(* IEC 61131-3 sources: s7-to-codesys/tests/POUs/ScenariosLang/FB_ConveyorStl_ScenarioTest, 15 files *)

(* ---- FB_ConveyorStl_ScenarioTest.decl.st ---- *)
// AUTO-GENERATED — не редактировать: s7conv gen-tests, сценарии scenarios/lang/FB_ConveyorStl.csv
// Правка — в CSV (scenarios/README.md), затем python -m s7conv build-corpus.
// Назначение: тесты поведения сконвертированного FB_ConveyorStl по сценариям CSV (сценариев: 7, строк: 58):
//             один метод-тест на сценарий, строки — по порядку с моделируемым временем GVL_S7Clock.
//             Ожидаемые значения — из CSV (эталонные модели по описанию логики блока), не из
//             результата конвертации.
// Автор:      s7conv 0.1.0 (сгенерировано)
// Версия:     не указана
// Документ:   scenarios/README.md, docs/methodology.md, раздел «Проверка поведения»
FUNCTION_BLOCK FB_ConveyorStl_ScenarioTest EXTENDS coUnit.FB_TestSuite
VAR
    fbStartSequence : FB_ConveyorStl;  // свой экземпляр на сценарий
    xStartSequenceDone : BOOL;  // сценарий выполнен (выполняется один раз)
    fbStopRunOut : FB_ConveyorStl;  // свой экземпляр на сценарий
    xStopRunOutDone : BOOL;  // сценарий выполнен (выполняется один раз)
    fbJamWithoutProducts : FB_ConveyorStl;  // свой экземпляр на сценарий
    xJamWithoutProductsDone : BOOL;  // сценарий выполнен (выполняется один раз)
    fbProductsKeepFlow : FB_ConveyorStl;  // свой экземпляр на сценарий
    xProductsKeepFlowDone : BOOL;  // сценарий выполнен (выполняется один раз)
    fbCountResetIsLevel : FB_ConveyorStl;  // свой экземпляр на сценарий
    xCountResetIsLevelDone : BOOL;  // сценарий выполнен (выполняется один раз)
    fbHornCutShort : FB_ConveyorStl;  // свой экземпляр на сценарий
    xHornCutShortDone : BOOL;  // сценарий выполнен (выполняется один раз)
    fbAckRestartsFlowWatch : FB_ConveyorStl;  // свой экземпляр на сценарий
    xAckRestartsFlowWatchDone : BOOL;  // сценарий выполнен (выполняется один раз)
END_VAR

(* ---- AckRestartsFlowWatch.method.decl.st ---- *)
// AUTO-GENERATED — не редактировать: scenarios/lang/FB_ConveyorStl.csv, сценарий AckRestartsFlowWatch (строк: 10)
METHOD PRIVATE AckRestartsFlowWatch
VAR
    stTimerZero : ST_S5Timer;  // пустое слово S5 для сброса
    stCounterZero : ST_S5Counter;  // пустое слово S5 для сброса
    iS5 : INT;  // номер таймера/счётчика S5
END_VAR

(* ---- AckRestartsFlowWatch.method.impl.st ---- *)
// AUTO-GENERATED — не редактировать: scenarios/lang/FB_ConveyorStl.csv, сценарий AckRestartsFlowWatch
coUnit.TEST('AckRestartsFlowWatch');
IF NOT xAckRestartsFlowWatchDone THEN
    xAckRestartsFlowWatchDone := TRUE;
    GVL_S7Clock.xSimulation := TRUE;
    // слова S5 — глобальные (GVL_S5Timers_Lang): сценарий начинается с чистых таймеров и счётчиков
    FOR iS5 := 0 TO 5 DO
        GVL_S5Timers_Lang.aTimer[iS5] := stTimerZero;
    END_FOR
    // слова S5 — глобальные (GVL_S5Counters_Lang): сценарий начинается с чистых таймеров и счётчиков
    FOR iS5 := 0 TO 1 DO
        GVL_S5Counters_Lang.aCounter[iS5] := stCounterZero;
    END_FOR

    // #1, t = 0 мс — пуск: запрос, сирена T1 и задержка T2 пошли
    GVL_S7Clock.tSimNow := T#0MS;
    fbAckRestartsFlowWatch.xStart := TRUE;
    fbAckRestartsFlowWatch.xStop := FALSE;
    fbAckRestartsFlowWatch.xSensor := FALSE;
    fbAckRestartsFlowWatch.xAck := FALSE;
    fbAckRestartsFlowWatch.xCountReset := FALSE;
    fbAckRestartsFlowWatch();
    AssertEquals_BOOL(Expected := TRUE,
                      Actual := fbAckRestartsFlowWatch.xHorn,
                      Message := 'AckRestartsFlowWatch#1 xHorn');
    AssertEquals_BOOL(Expected := FALSE,
                      Actual := fbAckRestartsFlowWatch.xMotor,
                      Message := 'AckRestartsFlowWatch#1 xMotor');
    AssertEquals_BOOL(Expected := FALSE,
                      Actual := fbAckRestartsFlowWatch.xFlowOk,
                      Message := 'AckRestartsFlowWatch#1 xFlowOk');
    AssertEquals_BOOL(Expected := FALSE,
                      Actual := fbAckRestartsFlowWatch.xJam,
                      Message := 'AckRestartsFlowWatch#1 xJam');
    AssertEquals_INT(Expected := 200,
                     Actual := fbAckRestartsFlowWatch.iDelayLeft,
                     Message := 'AckRestartsFlowWatch#1 iDelayLeft');
    AssertEquals_WORD(Expected := 16#0000,
                      Actual := fbAckRestartsFlowWatch.wRunOutBcd,
                      Message := 'AckRestartsFlowWatch#1 wRunOutBcd');
    AssertEquals_INT(Expected := 0,
                     Actual := fbAckRestartsFlowWatch.iCount,
                     Message := 'AckRestartsFlowWatch#1 iCount');
    AssertEquals_WORD(Expected := 16#0000,
                      Actual := fbAckRestartsFlowWatch.wCountBcd,
                      Message := 'AckRestartsFlowWatch#1 wCountBcd');

    // #2, t = 100 мс — кнопка отпущена
    GVL_S7Clock.tSimNow := T#100MS;
    fbAckRestartsFlowWatch.xStart := FALSE;
    fbAckRestartsFlowWatch();
    AssertEquals_BOOL(Expected := TRUE,
                      Actual := fbAckRestartsFlowWatch.xHorn,
                      Message := 'AckRestartsFlowWatch#2 xHorn');
    AssertEquals_BOOL(Expected := FALSE,
                      Actual := fbAckRestartsFlowWatch.xMotor,
                      Message := 'AckRestartsFlowWatch#2 xMotor');
    AssertEquals_BOOL(Expected := FALSE,
                      Actual := fbAckRestartsFlowWatch.xFlowOk,
                      Message := 'AckRestartsFlowWatch#2 xFlowOk');
    AssertEquals_BOOL(Expected := FALSE,
                      Actual := fbAckRestartsFlowWatch.xJam,
                      Message := 'AckRestartsFlowWatch#2 xJam');
    AssertEquals_INT(Expected := 190,
                     Actual := fbAckRestartsFlowWatch.iDelayLeft,
                     Message := 'AckRestartsFlowWatch#2 iDelayLeft');
    AssertEquals_WORD(Expected := 16#0000,
                      Actual := fbAckRestartsFlowWatch.wRunOutBcd,
                      Message := 'AckRestartsFlowWatch#2 wRunOutBcd');
    AssertEquals_INT(Expected := 0,
                     Actual := fbAckRestartsFlowWatch.iCount,
                     Message := 'AckRestartsFlowWatch#2 iCount');
    AssertEquals_WORD(Expected := 16#0000,
                      Actual := fbAckRestartsFlowWatch.wCountBcd,
                      Message := 'AckRestartsFlowWatch#2 wCountBcd');

    // #3, t = 2000 мс, на пороге таймера — 2 с: задержка T2 истекла — двигатель (T3 = 1)
    GVL_S7Clock.tSimNow := T#2000MS;
    fbAckRestartsFlowWatch();
    AssertEquals_BOOL(Expected := FALSE,
                      Actual := fbAckRestartsFlowWatch.xHorn,
                      Message := 'AckRestartsFlowWatch#3 xHorn');
    AssertEquals_BOOL(Expected := TRUE,
                      Actual := fbAckRestartsFlowWatch.xMotor,
                      Message := 'AckRestartsFlowWatch#3 xMotor');
    AssertEquals_BOOL(Expected := FALSE,
                      Actual := fbAckRestartsFlowWatch.xFlowOk,
                      Message := 'AckRestartsFlowWatch#3 xFlowOk');
    AssertEquals_BOOL(Expected := FALSE,
                      Actual := fbAckRestartsFlowWatch.xJam,
                      Message := 'AckRestartsFlowWatch#3 xJam');
    AssertEquals_INT(Expected := 0,
                     Actual := fbAckRestartsFlowWatch.iDelayLeft,
                     Message := 'AckRestartsFlowWatch#3 iDelayLeft');
    AssertEquals_WORD(Expected := 16#0000,
                      Actual := fbAckRestartsFlowWatch.wRunOutBcd,
                      Message := 'AckRestartsFlowWatch#3 wRunOutBcd');
    AssertEquals_INT(Expected := 0,
                     Actual := fbAckRestartsFlowWatch.iCount,
                     Message := 'AckRestartsFlowWatch#3 iCount');
    AssertEquals_WORD(Expected := 16#0000,
                      Actual := fbAckRestartsFlowWatch.wCountBcd,
                      Message := 'AckRestartsFlowWatch#3 wCountBcd');

    // #4, t = 2500 мс — датчик залип в 1: T4 пошёл один раз, изделие №1
    GVL_S7Clock.tSimNow := T#2500MS;
    fbAckRestartsFlowWatch.xSensor := TRUE;
    fbAckRestartsFlowWatch();
    AssertEquals_BOOL(Expected := FALSE,
                      Actual := fbAckRestartsFlowWatch.xHorn,
                      Message := 'AckRestartsFlowWatch#4 xHorn');
    AssertEquals_BOOL(Expected := TRUE,
                      Actual := fbAckRestartsFlowWatch.xMotor,
                      Message := 'AckRestartsFlowWatch#4 xMotor');
    AssertEquals_BOOL(Expected := TRUE,
                      Actual := fbAckRestartsFlowWatch.xFlowOk,
                      Message := 'AckRestartsFlowWatch#4 xFlowOk');
    AssertEquals_BOOL(Expected := FALSE,
                      Actual := fbAckRestartsFlowWatch.xJam,
                      Message := 'AckRestartsFlowWatch#4 xJam');
    AssertEquals_INT(Expected := 0,
                     Actual := fbAckRestartsFlowWatch.iDelayLeft,
                     Message := 'AckRestartsFlowWatch#4 iDelayLeft');
    AssertEquals_WORD(Expected := 16#0000,
                      Actual := fbAckRestartsFlowWatch.wRunOutBcd,
                      Message := 'AckRestartsFlowWatch#4 wRunOutBcd');
    AssertEquals_INT(Expected := 1,
                     Actual := fbAckRestartsFlowWatch.iCount,
                     Message := 'AckRestartsFlowWatch#4 iCount');
    AssertEquals_WORD(Expected := 16#0001,
                      Actual := fbAckRestartsFlowWatch.wCountBcd,
                      Message := 'AckRestartsFlowWatch#4 wCountBcd');

    // #5, t = 6500 мс, на пороге таймера — 4 с: T4 истёк, фронтов нет
    GVL_S7Clock.tSimNow := T#6500MS;
    fbAckRestartsFlowWatch();
    AssertEquals_BOOL(Expected := FALSE,
                      Actual := fbAckRestartsFlowWatch.xHorn,
                      Message := 'AckRestartsFlowWatch#5 xHorn');
    AssertEquals_BOOL(Expected := TRUE,
                      Actual := fbAckRestartsFlowWatch.xMotor,
                      Message := 'AckRestartsFlowWatch#5 xMotor');
    AssertEquals_BOOL(Expected := FALSE,
                      Actual := fbAckRestartsFlowWatch.xFlowOk,
                      Message := 'AckRestartsFlowWatch#5 xFlowOk');
    AssertEquals_BOOL(Expected := FALSE,
                      Actual := fbAckRestartsFlowWatch.xJam,
                      Message := 'AckRestartsFlowWatch#5 xJam');
    AssertEquals_INT(Expected := 0,
                     Actual := fbAckRestartsFlowWatch.iDelayLeft,
                     Message := 'AckRestartsFlowWatch#5 iDelayLeft');
    AssertEquals_WORD(Expected := 16#0000,
                      Actual := fbAckRestartsFlowWatch.wRunOutBcd,
                      Message := 'AckRestartsFlowWatch#5 wRunOutBcd');
    AssertEquals_INT(Expected := 1,
                     Actual := fbAckRestartsFlowWatch.iCount,
                     Message := 'AckRestartsFlowWatch#5 iCount');
    AssertEquals_WORD(Expected := 16#0001,
                      Actual := fbAckRestartsFlowWatch.wCountBcd,
                      Message := 'AckRestartsFlowWatch#5 wCountBcd');

    // #6, t = 7000 мс, на пороге таймера — контроль взведён: затор
    GVL_S7Clock.tSimNow := T#7000MS;
    fbAckRestartsFlowWatch();
    AssertEquals_BOOL(Expected := FALSE,
                      Actual := fbAckRestartsFlowWatch.xHorn,
                      Message := 'AckRestartsFlowWatch#6 xHorn');
    AssertEquals_BOOL(Expected := TRUE,
                      Actual := fbAckRestartsFlowWatch.xMotor,
                      Message := 'AckRestartsFlowWatch#6 xMotor');
    AssertEquals_BOOL(Expected := FALSE,
                      Actual := fbAckRestartsFlowWatch.xFlowOk,
                      Message := 'AckRestartsFlowWatch#6 xFlowOk');
    AssertEquals_BOOL(Expected := TRUE,
                      Actual := fbAckRestartsFlowWatch.xJam,
                      Message := 'AckRestartsFlowWatch#6 xJam');
    AssertEquals_INT(Expected := 0,
                     Actual := fbAckRestartsFlowWatch.iDelayLeft,
                     Message := 'AckRestartsFlowWatch#6 iDelayLeft');
    AssertEquals_WORD(Expected := 16#0000,
                      Actual := fbAckRestartsFlowWatch.wRunOutBcd,
                      Message := 'AckRestartsFlowWatch#6 wRunOutBcd');
    AssertEquals_INT(Expected := 1,
                     Actual := fbAckRestartsFlowWatch.iCount,
                     Message := 'AckRestartsFlowWatch#6 iCount');
    AssertEquals_WORD(Expected := 16#0001,
                      Actual := fbAckRestartsFlowWatch.wCountBcd,
                      Message := 'AckRestartsFlowWatch#6 wCountBcd');

    // #7, t = 7100 мс — запрос снят: выбег
    GVL_S7Clock.tSimNow := T#7100MS;
    fbAckRestartsFlowWatch();
    AssertEquals_BOOL(Expected := FALSE,
                      Actual := fbAckRestartsFlowWatch.xHorn,
                      Message := 'AckRestartsFlowWatch#7 xHorn');
    AssertEquals_BOOL(Expected := TRUE,
                      Actual := fbAckRestartsFlowWatch.xMotor,
                      Message := 'AckRestartsFlowWatch#7 xMotor');
    AssertEquals_BOOL(Expected := FALSE,
                      Actual := fbAckRestartsFlowWatch.xFlowOk,
                      Message := 'AckRestartsFlowWatch#7 xFlowOk');
    AssertEquals_BOOL(Expected := TRUE,
                      Actual := fbAckRestartsFlowWatch.xJam,
                      Message := 'AckRestartsFlowWatch#7 xJam');
    AssertEquals_INT(Expected := 0,
                     Actual := fbAckRestartsFlowWatch.iDelayLeft,
                     Message := 'AckRestartsFlowWatch#7 iDelayLeft');
    AssertEquals_WORD(Expected := 16#0300,
                      Actual := fbAckRestartsFlowWatch.wRunOutBcd,
                      Message := 'AckRestartsFlowWatch#7 wRunOutBcd');
    AssertEquals_INT(Expected := 1,
                     Actual := fbAckRestartsFlowWatch.iCount,
                     Message := 'AckRestartsFlowWatch#7 iCount');
    AssertEquals_WORD(Expected := 16#0001,
                      Actual := fbAckRestartsFlowWatch.wCountBcd,
                      Message := 'AckRestartsFlowWatch#7 wCountBcd');

    // #8, t = 10100 мс, на пороге таймера — выбег закончен
    GVL_S7Clock.tSimNow := T#10100MS;
    fbAckRestartsFlowWatch();
    AssertEquals_BOOL(Expected := FALSE,
                      Actual := fbAckRestartsFlowWatch.xHorn,
                      Message := 'AckRestartsFlowWatch#8 xHorn');
    AssertEquals_BOOL(Expected := FALSE,
                      Actual := fbAckRestartsFlowWatch.xMotor,
                      Message := 'AckRestartsFlowWatch#8 xMotor');
    AssertEquals_BOOL(Expected := FALSE,
                      Actual := fbAckRestartsFlowWatch.xFlowOk,
                      Message := 'AckRestartsFlowWatch#8 xFlowOk');
    AssertEquals_BOOL(Expected := TRUE,
                      Actual := fbAckRestartsFlowWatch.xJam,
                      Message := 'AckRestartsFlowWatch#8 xJam');
    AssertEquals_INT(Expected := 0,
                     Actual := fbAckRestartsFlowWatch.iDelayLeft,
                     Message := 'AckRestartsFlowWatch#8 iDelayLeft');
    AssertEquals_WORD(Expected := 16#0000,
                      Actual := fbAckRestartsFlowWatch.wRunOutBcd,
                      Message := 'AckRestartsFlowWatch#8 wRunOutBcd');
    AssertEquals_INT(Expected := 1,
                     Actual := fbAckRestartsFlowWatch.iCount,
                     Message := 'AckRestartsFlowWatch#8 iCount');
    AssertEquals_WORD(Expected := 16#0001,
                      Actual := fbAckRestartsFlowWatch.wCountBcd,
                      Message := 'AckRestartsFlowWatch#8 wCountBcd');

    // #9, t = 10500 мс — квитирование: затор снят, FR T4 (SE в этом вызове уже прошёл)
    GVL_S7Clock.tSimNow := T#10500MS;
    fbAckRestartsFlowWatch.xAck := TRUE;
    fbAckRestartsFlowWatch();
    AssertEquals_BOOL(Expected := FALSE,
                      Actual := fbAckRestartsFlowWatch.xHorn,
                      Message := 'AckRestartsFlowWatch#9 xHorn');
    AssertEquals_BOOL(Expected := FALSE,
                      Actual := fbAckRestartsFlowWatch.xMotor,
                      Message := 'AckRestartsFlowWatch#9 xMotor');
    AssertEquals_BOOL(Expected := FALSE,
                      Actual := fbAckRestartsFlowWatch.xFlowOk,
                      Message := 'AckRestartsFlowWatch#9 xFlowOk');
    AssertEquals_BOOL(Expected := FALSE,
                      Actual := fbAckRestartsFlowWatch.xJam,
                      Message := 'AckRestartsFlowWatch#9 xJam');
    AssertEquals_INT(Expected := 0,
                     Actual := fbAckRestartsFlowWatch.iDelayLeft,
                     Message := 'AckRestartsFlowWatch#9 iDelayLeft');
    AssertEquals_WORD(Expected := 16#0000,
                      Actual := fbAckRestartsFlowWatch.wRunOutBcd,
                      Message := 'AckRestartsFlowWatch#9 wRunOutBcd');
    AssertEquals_INT(Expected := 1,
                     Actual := fbAckRestartsFlowWatch.iCount,
                     Message := 'AckRestartsFlowWatch#9 iCount');
    AssertEquals_WORD(Expected := 16#0001,
                      Actual := fbAckRestartsFlowWatch.wCountBcd,
                      Message := 'AckRestartsFlowWatch#9 wCountBcd');

    // #10, t = 10600 мс — следующий вызов: SE видит фронт — T4 перезапущен
    GVL_S7Clock.tSimNow := T#10600MS;
    fbAckRestartsFlowWatch.xAck := FALSE;
    fbAckRestartsFlowWatch();
    AssertEquals_BOOL(Expected := FALSE,
                      Actual := fbAckRestartsFlowWatch.xHorn,
                      Message := 'AckRestartsFlowWatch#10 xHorn');
    AssertEquals_BOOL(Expected := FALSE,
                      Actual := fbAckRestartsFlowWatch.xMotor,
                      Message := 'AckRestartsFlowWatch#10 xMotor');
    AssertEquals_BOOL(Expected := TRUE,
                      Actual := fbAckRestartsFlowWatch.xFlowOk,
                      Message := 'AckRestartsFlowWatch#10 xFlowOk');
    AssertEquals_BOOL(Expected := FALSE,
                      Actual := fbAckRestartsFlowWatch.xJam,
                      Message := 'AckRestartsFlowWatch#10 xJam');
    AssertEquals_INT(Expected := 0,
                     Actual := fbAckRestartsFlowWatch.iDelayLeft,
                     Message := 'AckRestartsFlowWatch#10 iDelayLeft');
    AssertEquals_WORD(Expected := 16#0000,
                      Actual := fbAckRestartsFlowWatch.wRunOutBcd,
                      Message := 'AckRestartsFlowWatch#10 wRunOutBcd');
    AssertEquals_INT(Expected := 1,
                     Actual := fbAckRestartsFlowWatch.iCount,
                     Message := 'AckRestartsFlowWatch#10 iCount');
    AssertEquals_WORD(Expected := 16#0001,
                      Actual := fbAckRestartsFlowWatch.wCountBcd,
                      Message := 'AckRestartsFlowWatch#10 wCountBcd');

    GVL_S7Clock.xSimulation := FALSE;
END_IF
coUnit.TEST_FINISHED();

(* ---- CountResetIsLevel.method.decl.st ---- *)
// AUTO-GENERATED — не редактировать: scenarios/lang/FB_ConveyorStl.csv, сценарий CountResetIsLevel (строк: 8)
METHOD PRIVATE CountResetIsLevel
VAR
    stTimerZero : ST_S5Timer;  // пустое слово S5 для сброса
    stCounterZero : ST_S5Counter;  // пустое слово S5 для сброса
    iS5 : INT;  // номер таймера/счётчика S5
END_VAR

(* ---- CountResetIsLevel.method.impl.st ---- *)
// AUTO-GENERATED — не редактировать: scenarios/lang/FB_ConveyorStl.csv, сценарий CountResetIsLevel
coUnit.TEST('CountResetIsLevel');
IF NOT xCountResetIsLevelDone THEN
    xCountResetIsLevelDone := TRUE;
    GVL_S7Clock.xSimulation := TRUE;
    // слова S5 — глобальные (GVL_S5Timers_Lang): сценарий начинается с чистых таймеров и счётчиков
    FOR iS5 := 0 TO 5 DO
        GVL_S5Timers_Lang.aTimer[iS5] := stTimerZero;
    END_FOR
    // слова S5 — глобальные (GVL_S5Counters_Lang): сценарий начинается с чистых таймеров и счётчиков
    FOR iS5 := 0 TO 1 DO
        GVL_S5Counters_Lang.aCounter[iS5] := stCounterZero;
    END_FOR

    // #1, t = 0 мс — изделие №1
    GVL_S7Clock.tSimNow := T#0MS;
    fbCountResetIsLevel.xStart := FALSE;
    fbCountResetIsLevel.xStop := FALSE;
    fbCountResetIsLevel.xSensor := TRUE;
    fbCountResetIsLevel.xAck := FALSE;
    fbCountResetIsLevel.xCountReset := FALSE;
    fbCountResetIsLevel();
    AssertEquals_BOOL(Expected := FALSE, Actual := fbCountResetIsLevel.xHorn, Message := 'CountResetIsLevel#1 xHorn');
    AssertEquals_BOOL(Expected := FALSE, Actual := fbCountResetIsLevel.xMotor, Message := 'CountResetIsLevel#1 xMotor');
    AssertEquals_BOOL(Expected := TRUE,
                      Actual := fbCountResetIsLevel.xFlowOk,
                      Message := 'CountResetIsLevel#1 xFlowOk');
    AssertEquals_BOOL(Expected := FALSE, Actual := fbCountResetIsLevel.xJam, Message := 'CountResetIsLevel#1 xJam');
    AssertEquals_INT(Expected := 0,
                     Actual := fbCountResetIsLevel.iDelayLeft,
                     Message := 'CountResetIsLevel#1 iDelayLeft');
    AssertEquals_WORD(Expected := 16#0000,
                      Actual := fbCountResetIsLevel.wRunOutBcd,
                      Message := 'CountResetIsLevel#1 wRunOutBcd');
    AssertEquals_INT(Expected := 1, Actual := fbCountResetIsLevel.iCount, Message := 'CountResetIsLevel#1 iCount');
    AssertEquals_WORD(Expected := 16#0001,
                      Actual := fbCountResetIsLevel.wCountBcd,
                      Message := 'CountResetIsLevel#1 wCountBcd');

    // #2, t = 100 мс — датчик свободен
    GVL_S7Clock.tSimNow := T#100MS;
    fbCountResetIsLevel.xSensor := FALSE;
    fbCountResetIsLevel();
    AssertEquals_BOOL(Expected := FALSE, Actual := fbCountResetIsLevel.xHorn, Message := 'CountResetIsLevel#2 xHorn');
    AssertEquals_BOOL(Expected := FALSE, Actual := fbCountResetIsLevel.xMotor, Message := 'CountResetIsLevel#2 xMotor');
    AssertEquals_BOOL(Expected := TRUE,
                      Actual := fbCountResetIsLevel.xFlowOk,
                      Message := 'CountResetIsLevel#2 xFlowOk');
    AssertEquals_BOOL(Expected := FALSE, Actual := fbCountResetIsLevel.xJam, Message := 'CountResetIsLevel#2 xJam');
    AssertEquals_INT(Expected := 0,
                     Actual := fbCountResetIsLevel.iDelayLeft,
                     Message := 'CountResetIsLevel#2 iDelayLeft');
    AssertEquals_WORD(Expected := 16#0000,
                      Actual := fbCountResetIsLevel.wRunOutBcd,
                      Message := 'CountResetIsLevel#2 wRunOutBcd');
    AssertEquals_INT(Expected := 1, Actual := fbCountResetIsLevel.iCount, Message := 'CountResetIsLevel#2 iCount');
    AssertEquals_WORD(Expected := 16#0001,
                      Actual := fbCountResetIsLevel.wCountBcd,
                      Message := 'CountResetIsLevel#2 wCountBcd');

    // #3, t = 200 мс — изделие №2
    GVL_S7Clock.tSimNow := T#200MS;
    fbCountResetIsLevel.xSensor := TRUE;
    fbCountResetIsLevel();
    AssertEquals_BOOL(Expected := FALSE, Actual := fbCountResetIsLevel.xHorn, Message := 'CountResetIsLevel#3 xHorn');
    AssertEquals_BOOL(Expected := FALSE, Actual := fbCountResetIsLevel.xMotor, Message := 'CountResetIsLevel#3 xMotor');
    AssertEquals_BOOL(Expected := TRUE,
                      Actual := fbCountResetIsLevel.xFlowOk,
                      Message := 'CountResetIsLevel#3 xFlowOk');
    AssertEquals_BOOL(Expected := FALSE, Actual := fbCountResetIsLevel.xJam, Message := 'CountResetIsLevel#3 xJam');
    AssertEquals_INT(Expected := 0,
                     Actual := fbCountResetIsLevel.iDelayLeft,
                     Message := 'CountResetIsLevel#3 iDelayLeft');
    AssertEquals_WORD(Expected := 16#0000,
                      Actual := fbCountResetIsLevel.wRunOutBcd,
                      Message := 'CountResetIsLevel#3 wRunOutBcd');
    AssertEquals_INT(Expected := 2, Actual := fbCountResetIsLevel.iCount, Message := 'CountResetIsLevel#3 iCount');
    AssertEquals_WORD(Expected := 16#0002,
                      Actual := fbCountResetIsLevel.wCountBcd,
                      Message := 'CountResetIsLevel#3 wCountBcd');

    // #4, t = 300 мс — датчик свободен
    GVL_S7Clock.tSimNow := T#300MS;
    fbCountResetIsLevel.xSensor := FALSE;
    fbCountResetIsLevel();
    AssertEquals_BOOL(Expected := FALSE, Actual := fbCountResetIsLevel.xHorn, Message := 'CountResetIsLevel#4 xHorn');
    AssertEquals_BOOL(Expected := FALSE, Actual := fbCountResetIsLevel.xMotor, Message := 'CountResetIsLevel#4 xMotor');
    AssertEquals_BOOL(Expected := TRUE,
                      Actual := fbCountResetIsLevel.xFlowOk,
                      Message := 'CountResetIsLevel#4 xFlowOk');
    AssertEquals_BOOL(Expected := FALSE, Actual := fbCountResetIsLevel.xJam, Message := 'CountResetIsLevel#4 xJam');
    AssertEquals_INT(Expected := 0,
                     Actual := fbCountResetIsLevel.iDelayLeft,
                     Message := 'CountResetIsLevel#4 iDelayLeft');
    AssertEquals_WORD(Expected := 16#0000,
                      Actual := fbCountResetIsLevel.wRunOutBcd,
                      Message := 'CountResetIsLevel#4 wRunOutBcd');
    AssertEquals_INT(Expected := 2, Actual := fbCountResetIsLevel.iCount, Message := 'CountResetIsLevel#4 iCount');
    AssertEquals_WORD(Expected := 16#0002,
                      Actual := fbCountResetIsLevel.wCountBcd,
                      Message := 'CountResetIsLevel#4 wCountBcd');

    // #5, t = 400 мс — сброс счётчика
    GVL_S7Clock.tSimNow := T#400MS;
    fbCountResetIsLevel.xCountReset := TRUE;
    fbCountResetIsLevel();
    AssertEquals_BOOL(Expected := FALSE, Actual := fbCountResetIsLevel.xHorn, Message := 'CountResetIsLevel#5 xHorn');
    AssertEquals_BOOL(Expected := FALSE, Actual := fbCountResetIsLevel.xMotor, Message := 'CountResetIsLevel#5 xMotor');
    AssertEquals_BOOL(Expected := TRUE,
                      Actual := fbCountResetIsLevel.xFlowOk,
                      Message := 'CountResetIsLevel#5 xFlowOk');
    AssertEquals_BOOL(Expected := FALSE, Actual := fbCountResetIsLevel.xJam, Message := 'CountResetIsLevel#5 xJam');
    AssertEquals_INT(Expected := 0,
                     Actual := fbCountResetIsLevel.iDelayLeft,
                     Message := 'CountResetIsLevel#5 iDelayLeft');
    AssertEquals_WORD(Expected := 16#0000,
                      Actual := fbCountResetIsLevel.wRunOutBcd,
                      Message := 'CountResetIsLevel#5 wRunOutBcd');
    AssertEquals_INT(Expected := 0, Actual := fbCountResetIsLevel.iCount, Message := 'CountResetIsLevel#5 iCount');
    AssertEquals_WORD(Expected := 16#0000,
                      Actual := fbCountResetIsLevel.wCountBcd,
                      Message := 'CountResetIsLevel#5 wCountBcd');

    // #6, t = 500 мс — изделие при нажатом сбросе: CU считает, R тут же обнуляет
    GVL_S7Clock.tSimNow := T#500MS;
    fbCountResetIsLevel.xSensor := TRUE;
    fbCountResetIsLevel();
    AssertEquals_BOOL(Expected := FALSE, Actual := fbCountResetIsLevel.xHorn, Message := 'CountResetIsLevel#6 xHorn');
    AssertEquals_BOOL(Expected := FALSE, Actual := fbCountResetIsLevel.xMotor, Message := 'CountResetIsLevel#6 xMotor');
    AssertEquals_BOOL(Expected := TRUE,
                      Actual := fbCountResetIsLevel.xFlowOk,
                      Message := 'CountResetIsLevel#6 xFlowOk');
    AssertEquals_BOOL(Expected := FALSE, Actual := fbCountResetIsLevel.xJam, Message := 'CountResetIsLevel#6 xJam');
    AssertEquals_INT(Expected := 0,
                     Actual := fbCountResetIsLevel.iDelayLeft,
                     Message := 'CountResetIsLevel#6 iDelayLeft');
    AssertEquals_WORD(Expected := 16#0000,
                      Actual := fbCountResetIsLevel.wRunOutBcd,
                      Message := 'CountResetIsLevel#6 wRunOutBcd');
    AssertEquals_INT(Expected := 0, Actual := fbCountResetIsLevel.iCount, Message := 'CountResetIsLevel#6 iCount');
    AssertEquals_WORD(Expected := 16#0000,
                      Actual := fbCountResetIsLevel.wCountBcd,
                      Message := 'CountResetIsLevel#6 wCountBcd');

    // #7, t = 600 мс — сброс отпущен
    GVL_S7Clock.tSimNow := T#600MS;
    fbCountResetIsLevel.xSensor := FALSE;
    fbCountResetIsLevel.xCountReset := FALSE;
    fbCountResetIsLevel();
    AssertEquals_BOOL(Expected := FALSE, Actual := fbCountResetIsLevel.xHorn, Message := 'CountResetIsLevel#7 xHorn');
    AssertEquals_BOOL(Expected := FALSE, Actual := fbCountResetIsLevel.xMotor, Message := 'CountResetIsLevel#7 xMotor');
    AssertEquals_BOOL(Expected := TRUE,
                      Actual := fbCountResetIsLevel.xFlowOk,
                      Message := 'CountResetIsLevel#7 xFlowOk');
    AssertEquals_BOOL(Expected := FALSE, Actual := fbCountResetIsLevel.xJam, Message := 'CountResetIsLevel#7 xJam');
    AssertEquals_INT(Expected := 0,
                     Actual := fbCountResetIsLevel.iDelayLeft,
                     Message := 'CountResetIsLevel#7 iDelayLeft');
    AssertEquals_WORD(Expected := 16#0000,
                      Actual := fbCountResetIsLevel.wRunOutBcd,
                      Message := 'CountResetIsLevel#7 wRunOutBcd');
    AssertEquals_INT(Expected := 0, Actual := fbCountResetIsLevel.iCount, Message := 'CountResetIsLevel#7 iCount');
    AssertEquals_WORD(Expected := 16#0000,
                      Actual := fbCountResetIsLevel.wCountBcd,
                      Message := 'CountResetIsLevel#7 wCountBcd');

    // #8, t = 700 мс — изделие №1 после сброса
    GVL_S7Clock.tSimNow := T#700MS;
    fbCountResetIsLevel.xSensor := TRUE;
    fbCountResetIsLevel();
    AssertEquals_BOOL(Expected := FALSE, Actual := fbCountResetIsLevel.xHorn, Message := 'CountResetIsLevel#8 xHorn');
    AssertEquals_BOOL(Expected := FALSE, Actual := fbCountResetIsLevel.xMotor, Message := 'CountResetIsLevel#8 xMotor');
    AssertEquals_BOOL(Expected := TRUE,
                      Actual := fbCountResetIsLevel.xFlowOk,
                      Message := 'CountResetIsLevel#8 xFlowOk');
    AssertEquals_BOOL(Expected := FALSE, Actual := fbCountResetIsLevel.xJam, Message := 'CountResetIsLevel#8 xJam');
    AssertEquals_INT(Expected := 0,
                     Actual := fbCountResetIsLevel.iDelayLeft,
                     Message := 'CountResetIsLevel#8 iDelayLeft');
    AssertEquals_WORD(Expected := 16#0000,
                      Actual := fbCountResetIsLevel.wRunOutBcd,
                      Message := 'CountResetIsLevel#8 wRunOutBcd');
    AssertEquals_INT(Expected := 1, Actual := fbCountResetIsLevel.iCount, Message := 'CountResetIsLevel#8 iCount');
    AssertEquals_WORD(Expected := 16#0001,
                      Actual := fbCountResetIsLevel.wCountBcd,
                      Message := 'CountResetIsLevel#8 wCountBcd');

    GVL_S7Clock.xSimulation := FALSE;
END_IF
coUnit.TEST_FINISHED();

(* ---- HornCutShort.method.decl.st ---- *)
// AUTO-GENERATED — не редактировать: scenarios/lang/FB_ConveyorStl.csv, сценарий HornCutShort (строк: 4)
METHOD PRIVATE HornCutShort
VAR
    stTimerZero : ST_S5Timer;  // пустое слово S5 для сброса
    stCounterZero : ST_S5Counter;  // пустое слово S5 для сброса
    iS5 : INT;  // номер таймера/счётчика S5
END_VAR

(* ---- HornCutShort.method.impl.st ---- *)
// AUTO-GENERATED — не редактировать: scenarios/lang/FB_ConveyorStl.csv, сценарий HornCutShort
coUnit.TEST('HornCutShort');
IF NOT xHornCutShortDone THEN
    xHornCutShortDone := TRUE;
    GVL_S7Clock.xSimulation := TRUE;
    // слова S5 — глобальные (GVL_S5Timers_Lang): сценарий начинается с чистых таймеров и счётчиков
    FOR iS5 := 0 TO 5 DO
        GVL_S5Timers_Lang.aTimer[iS5] := stTimerZero;
    END_FOR
    // слова S5 — глобальные (GVL_S5Counters_Lang): сценарий начинается с чистых таймеров и счётчиков
    FOR iS5 := 0 TO 1 DO
        GVL_S5Counters_Lang.aCounter[iS5] := stCounterZero;
    END_FOR

    // #1, t = 0 мс — пуск: сирена, остаток 200
    GVL_S7Clock.tSimNow := T#0MS;
    fbHornCutShort.xStart := TRUE;
    fbHornCutShort.xStop := FALSE;
    fbHornCutShort.xSensor := FALSE;
    fbHornCutShort.xAck := FALSE;
    fbHornCutShort.xCountReset := FALSE;
    fbHornCutShort();
    AssertEquals_BOOL(Expected := TRUE, Actual := fbHornCutShort.xHorn, Message := 'HornCutShort#1 xHorn');
    AssertEquals_BOOL(Expected := FALSE, Actual := fbHornCutShort.xMotor, Message := 'HornCutShort#1 xMotor');
    AssertEquals_BOOL(Expected := FALSE, Actual := fbHornCutShort.xFlowOk, Message := 'HornCutShort#1 xFlowOk');
    AssertEquals_BOOL(Expected := FALSE, Actual := fbHornCutShort.xJam, Message := 'HornCutShort#1 xJam');
    AssertEquals_INT(Expected := 200, Actual := fbHornCutShort.iDelayLeft, Message := 'HornCutShort#1 iDelayLeft');
    AssertEquals_WORD(Expected := 16#0000, Actual := fbHornCutShort.wRunOutBcd, Message := 'HornCutShort#1 wRunOutBcd');
    AssertEquals_INT(Expected := 0, Actual := fbHornCutShort.iCount, Message := 'HornCutShort#1 iCount');
    AssertEquals_WORD(Expected := 16#0000, Actual := fbHornCutShort.wCountBcd, Message := 'HornCutShort#1 wCountBcd');

    // #2, t = 300 мс — стоп: сирена оборвана, T2 остановлен с остатком 170
    GVL_S7Clock.tSimNow := T#300MS;
    fbHornCutShort.xStart := FALSE;
    fbHornCutShort.xStop := TRUE;
    fbHornCutShort();
    AssertEquals_BOOL(Expected := FALSE, Actual := fbHornCutShort.xHorn, Message := 'HornCutShort#2 xHorn');
    AssertEquals_BOOL(Expected := FALSE, Actual := fbHornCutShort.xMotor, Message := 'HornCutShort#2 xMotor');
    AssertEquals_BOOL(Expected := FALSE, Actual := fbHornCutShort.xFlowOk, Message := 'HornCutShort#2 xFlowOk');
    AssertEquals_BOOL(Expected := FALSE, Actual := fbHornCutShort.xJam, Message := 'HornCutShort#2 xJam');
    AssertEquals_INT(Expected := 170, Actual := fbHornCutShort.iDelayLeft, Message := 'HornCutShort#2 iDelayLeft');
    AssertEquals_WORD(Expected := 16#0000, Actual := fbHornCutShort.wRunOutBcd, Message := 'HornCutShort#2 wRunOutBcd');
    AssertEquals_INT(Expected := 0, Actual := fbHornCutShort.iCount, Message := 'HornCutShort#2 iCount');
    AssertEquals_WORD(Expected := 16#0000, Actual := fbHornCutShort.wCountBcd, Message := 'HornCutShort#2 wCountBcd');

    // #3, t = 400 мс — остаток 170 сохраняется
    GVL_S7Clock.tSimNow := T#400MS;
    fbHornCutShort.xStop := FALSE;
    fbHornCutShort();
    AssertEquals_BOOL(Expected := FALSE, Actual := fbHornCutShort.xHorn, Message := 'HornCutShort#3 xHorn');
    AssertEquals_BOOL(Expected := FALSE, Actual := fbHornCutShort.xMotor, Message := 'HornCutShort#3 xMotor');
    AssertEquals_BOOL(Expected := FALSE, Actual := fbHornCutShort.xFlowOk, Message := 'HornCutShort#3 xFlowOk');
    AssertEquals_BOOL(Expected := FALSE, Actual := fbHornCutShort.xJam, Message := 'HornCutShort#3 xJam');
    AssertEquals_INT(Expected := 170, Actual := fbHornCutShort.iDelayLeft, Message := 'HornCutShort#3 iDelayLeft');
    AssertEquals_WORD(Expected := 16#0000, Actual := fbHornCutShort.wRunOutBcd, Message := 'HornCutShort#3 wRunOutBcd');
    AssertEquals_INT(Expected := 0, Actual := fbHornCutShort.iCount, Message := 'HornCutShort#3 iCount');
    AssertEquals_WORD(Expected := 16#0000, Actual := fbHornCutShort.wCountBcd, Message := 'HornCutShort#3 wCountBcd');

    // #4, t = 5000 мс — остаток 170 сохраняется
    GVL_S7Clock.tSimNow := T#5000MS;
    fbHornCutShort();
    AssertEquals_BOOL(Expected := FALSE, Actual := fbHornCutShort.xHorn, Message := 'HornCutShort#4 xHorn');
    AssertEquals_BOOL(Expected := FALSE, Actual := fbHornCutShort.xMotor, Message := 'HornCutShort#4 xMotor');
    AssertEquals_BOOL(Expected := FALSE, Actual := fbHornCutShort.xFlowOk, Message := 'HornCutShort#4 xFlowOk');
    AssertEquals_BOOL(Expected := FALSE, Actual := fbHornCutShort.xJam, Message := 'HornCutShort#4 xJam');
    AssertEquals_INT(Expected := 170, Actual := fbHornCutShort.iDelayLeft, Message := 'HornCutShort#4 iDelayLeft');
    AssertEquals_WORD(Expected := 16#0000, Actual := fbHornCutShort.wRunOutBcd, Message := 'HornCutShort#4 wRunOutBcd');
    AssertEquals_INT(Expected := 0, Actual := fbHornCutShort.iCount, Message := 'HornCutShort#4 iCount');
    AssertEquals_WORD(Expected := 16#0000, Actual := fbHornCutShort.wCountBcd, Message := 'HornCutShort#4 wCountBcd');

    GVL_S7Clock.xSimulation := FALSE;
END_IF
coUnit.TEST_FINISHED();

(* ---- JamWithoutProducts.method.decl.st ---- *)
// AUTO-GENERATED — не редактировать: scenarios/lang/FB_ConveyorStl.csv, сценарий JamWithoutProducts (строк: 9)
METHOD PRIVATE JamWithoutProducts
VAR
    stTimerZero : ST_S5Timer;  // пустое слово S5 для сброса
    stCounterZero : ST_S5Counter;  // пустое слово S5 для сброса
    iS5 : INT;  // номер таймера/счётчика S5
END_VAR

(* ---- JamWithoutProducts.method.impl.st ---- *)
// AUTO-GENERATED — не редактировать: scenarios/lang/FB_ConveyorStl.csv, сценарий JamWithoutProducts
coUnit.TEST('JamWithoutProducts');
IF NOT xJamWithoutProductsDone THEN
    xJamWithoutProductsDone := TRUE;
    GVL_S7Clock.xSimulation := TRUE;
    // слова S5 — глобальные (GVL_S5Timers_Lang): сценарий начинается с чистых таймеров и счётчиков
    FOR iS5 := 0 TO 5 DO
        GVL_S5Timers_Lang.aTimer[iS5] := stTimerZero;
    END_FOR
    // слова S5 — глобальные (GVL_S5Counters_Lang): сценарий начинается с чистых таймеров и счётчиков
    FOR iS5 := 0 TO 1 DO
        GVL_S5Counters_Lang.aCounter[iS5] := stCounterZero;
    END_FOR

    // #1, t = 0 мс — пуск: запрос, сирена T1 и задержка T2 пошли
    GVL_S7Clock.tSimNow := T#0MS;
    fbJamWithoutProducts.xStart := TRUE;
    fbJamWithoutProducts.xStop := FALSE;
    fbJamWithoutProducts.xSensor := FALSE;
    fbJamWithoutProducts.xAck := FALSE;
    fbJamWithoutProducts.xCountReset := FALSE;
    fbJamWithoutProducts();
    AssertEquals_BOOL(Expected := TRUE, Actual := fbJamWithoutProducts.xHorn, Message := 'JamWithoutProducts#1 xHorn');
    AssertEquals_BOOL(Expected := FALSE,
                      Actual := fbJamWithoutProducts.xMotor,
                      Message := 'JamWithoutProducts#1 xMotor');
    AssertEquals_BOOL(Expected := FALSE,
                      Actual := fbJamWithoutProducts.xFlowOk,
                      Message := 'JamWithoutProducts#1 xFlowOk');
    AssertEquals_BOOL(Expected := FALSE, Actual := fbJamWithoutProducts.xJam, Message := 'JamWithoutProducts#1 xJam');
    AssertEquals_INT(Expected := 200,
                     Actual := fbJamWithoutProducts.iDelayLeft,
                     Message := 'JamWithoutProducts#1 iDelayLeft');
    AssertEquals_WORD(Expected := 16#0000,
                      Actual := fbJamWithoutProducts.wRunOutBcd,
                      Message := 'JamWithoutProducts#1 wRunOutBcd');
    AssertEquals_INT(Expected := 0, Actual := fbJamWithoutProducts.iCount, Message := 'JamWithoutProducts#1 iCount');
    AssertEquals_WORD(Expected := 16#0000,
                      Actual := fbJamWithoutProducts.wCountBcd,
                      Message := 'JamWithoutProducts#1 wCountBcd');

    // #2, t = 100 мс — кнопка отпущена
    GVL_S7Clock.tSimNow := T#100MS;
    fbJamWithoutProducts.xStart := FALSE;
    fbJamWithoutProducts();
    AssertEquals_BOOL(Expected := TRUE, Actual := fbJamWithoutProducts.xHorn, Message := 'JamWithoutProducts#2 xHorn');
    AssertEquals_BOOL(Expected := FALSE,
                      Actual := fbJamWithoutProducts.xMotor,
                      Message := 'JamWithoutProducts#2 xMotor');
    AssertEquals_BOOL(Expected := FALSE,
                      Actual := fbJamWithoutProducts.xFlowOk,
                      Message := 'JamWithoutProducts#2 xFlowOk');
    AssertEquals_BOOL(Expected := FALSE, Actual := fbJamWithoutProducts.xJam, Message := 'JamWithoutProducts#2 xJam');
    AssertEquals_INT(Expected := 190,
                     Actual := fbJamWithoutProducts.iDelayLeft,
                     Message := 'JamWithoutProducts#2 iDelayLeft');
    AssertEquals_WORD(Expected := 16#0000,
                      Actual := fbJamWithoutProducts.wRunOutBcd,
                      Message := 'JamWithoutProducts#2 wRunOutBcd');
    AssertEquals_INT(Expected := 0, Actual := fbJamWithoutProducts.iCount, Message := 'JamWithoutProducts#2 iCount');
    AssertEquals_WORD(Expected := 16#0000,
                      Actual := fbJamWithoutProducts.wCountBcd,
                      Message := 'JamWithoutProducts#2 wCountBcd');

    // #3, t = 2000 мс, на пороге таймера — 2 с: задержка T2 истекла — двигатель (T3 = 1)
    GVL_S7Clock.tSimNow := T#2000MS;
    fbJamWithoutProducts();
    AssertEquals_BOOL(Expected := FALSE, Actual := fbJamWithoutProducts.xHorn, Message := 'JamWithoutProducts#3 xHorn');
    AssertEquals_BOOL(Expected := TRUE,
                      Actual := fbJamWithoutProducts.xMotor,
                      Message := 'JamWithoutProducts#3 xMotor');
    AssertEquals_BOOL(Expected := FALSE,
                      Actual := fbJamWithoutProducts.xFlowOk,
                      Message := 'JamWithoutProducts#3 xFlowOk');
    AssertEquals_BOOL(Expected := FALSE, Actual := fbJamWithoutProducts.xJam, Message := 'JamWithoutProducts#3 xJam');
    AssertEquals_INT(Expected := 0,
                     Actual := fbJamWithoutProducts.iDelayLeft,
                     Message := 'JamWithoutProducts#3 iDelayLeft');
    AssertEquals_WORD(Expected := 16#0000,
                      Actual := fbJamWithoutProducts.wRunOutBcd,
                      Message := 'JamWithoutProducts#3 wRunOutBcd');
    AssertEquals_INT(Expected := 0, Actual := fbJamWithoutProducts.iCount, Message := 'JamWithoutProducts#3 iCount');
    AssertEquals_WORD(Expected := 16#0000,
                      Actual := fbJamWithoutProducts.wCountBcd,
                      Message := 'JamWithoutProducts#3 wCountBcd');

    // #4, t = 6700 мс — 4,7 с работы: контроль ещё не взведён
    GVL_S7Clock.tSimNow := T#6700MS;
    fbJamWithoutProducts();
    AssertEquals_BOOL(Expected := FALSE, Actual := fbJamWithoutProducts.xHorn, Message := 'JamWithoutProducts#4 xHorn');
    AssertEquals_BOOL(Expected := TRUE,
                      Actual := fbJamWithoutProducts.xMotor,
                      Message := 'JamWithoutProducts#4 xMotor');
    AssertEquals_BOOL(Expected := FALSE,
                      Actual := fbJamWithoutProducts.xFlowOk,
                      Message := 'JamWithoutProducts#4 xFlowOk');
    AssertEquals_BOOL(Expected := FALSE, Actual := fbJamWithoutProducts.xJam, Message := 'JamWithoutProducts#4 xJam');
    AssertEquals_INT(Expected := 0,
                     Actual := fbJamWithoutProducts.iDelayLeft,
                     Message := 'JamWithoutProducts#4 iDelayLeft');
    AssertEquals_WORD(Expected := 16#0000,
                      Actual := fbJamWithoutProducts.wRunOutBcd,
                      Message := 'JamWithoutProducts#4 wRunOutBcd');
    AssertEquals_INT(Expected := 0, Actual := fbJamWithoutProducts.iCount, Message := 'JamWithoutProducts#4 iCount');
    AssertEquals_WORD(Expected := 16#0000,
                      Actual := fbJamWithoutProducts.wCountBcd,
                      Message := 'JamWithoutProducts#4 wCountBcd');

    // #5, t = 7000 мс, на пороге таймера — 5 с работы: T5 взвёл контроль, T4 не идёт — затор
    GVL_S7Clock.tSimNow := T#7000MS;
    fbJamWithoutProducts();
    AssertEquals_BOOL(Expected := FALSE, Actual := fbJamWithoutProducts.xHorn, Message := 'JamWithoutProducts#5 xHorn');
    AssertEquals_BOOL(Expected := TRUE,
                      Actual := fbJamWithoutProducts.xMotor,
                      Message := 'JamWithoutProducts#5 xMotor');
    AssertEquals_BOOL(Expected := FALSE,
                      Actual := fbJamWithoutProducts.xFlowOk,
                      Message := 'JamWithoutProducts#5 xFlowOk');
    AssertEquals_BOOL(Expected := TRUE, Actual := fbJamWithoutProducts.xJam, Message := 'JamWithoutProducts#5 xJam');
    AssertEquals_INT(Expected := 0,
                     Actual := fbJamWithoutProducts.iDelayLeft,
                     Message := 'JamWithoutProducts#5 iDelayLeft');
    AssertEquals_WORD(Expected := 16#0000,
                      Actual := fbJamWithoutProducts.wRunOutBcd,
                      Message := 'JamWithoutProducts#5 wRunOutBcd');
    AssertEquals_INT(Expected := 0, Actual := fbJamWithoutProducts.iCount, Message := 'JamWithoutProducts#5 iCount');
    AssertEquals_WORD(Expected := 16#0000,
                      Actual := fbJamWithoutProducts.wCountBcd,
                      Message := 'JamWithoutProducts#5 wCountBcd');

    // #6, t = 7100 мс — затор сбросил запрос: выбег 3 с
    GVL_S7Clock.tSimNow := T#7100MS;
    fbJamWithoutProducts();
    AssertEquals_BOOL(Expected := FALSE, Actual := fbJamWithoutProducts.xHorn, Message := 'JamWithoutProducts#6 xHorn');
    AssertEquals_BOOL(Expected := TRUE,
                      Actual := fbJamWithoutProducts.xMotor,
                      Message := 'JamWithoutProducts#6 xMotor');
    AssertEquals_BOOL(Expected := FALSE,
                      Actual := fbJamWithoutProducts.xFlowOk,
                      Message := 'JamWithoutProducts#6 xFlowOk');
    AssertEquals_BOOL(Expected := TRUE, Actual := fbJamWithoutProducts.xJam, Message := 'JamWithoutProducts#6 xJam');
    AssertEquals_INT(Expected := 0,
                     Actual := fbJamWithoutProducts.iDelayLeft,
                     Message := 'JamWithoutProducts#6 iDelayLeft');
    AssertEquals_WORD(Expected := 16#0300,
                      Actual := fbJamWithoutProducts.wRunOutBcd,
                      Message := 'JamWithoutProducts#6 wRunOutBcd');
    AssertEquals_INT(Expected := 0, Actual := fbJamWithoutProducts.iCount, Message := 'JamWithoutProducts#6 iCount');
    AssertEquals_WORD(Expected := 16#0000,
                      Actual := fbJamWithoutProducts.wCountBcd,
                      Message := 'JamWithoutProducts#6 wCountBcd');

    // #7, t = 10100 мс, на пороге таймера — выбег закончен: двигатель остановлен, T5 сброшен
    GVL_S7Clock.tSimNow := T#10100MS;
    fbJamWithoutProducts();
    AssertEquals_BOOL(Expected := FALSE, Actual := fbJamWithoutProducts.xHorn, Message := 'JamWithoutProducts#7 xHorn');
    AssertEquals_BOOL(Expected := FALSE,
                      Actual := fbJamWithoutProducts.xMotor,
                      Message := 'JamWithoutProducts#7 xMotor');
    AssertEquals_BOOL(Expected := FALSE,
                      Actual := fbJamWithoutProducts.xFlowOk,
                      Message := 'JamWithoutProducts#7 xFlowOk');
    AssertEquals_BOOL(Expected := TRUE, Actual := fbJamWithoutProducts.xJam, Message := 'JamWithoutProducts#7 xJam');
    AssertEquals_INT(Expected := 0,
                     Actual := fbJamWithoutProducts.iDelayLeft,
                     Message := 'JamWithoutProducts#7 iDelayLeft');
    AssertEquals_WORD(Expected := 16#0000,
                      Actual := fbJamWithoutProducts.wRunOutBcd,
                      Message := 'JamWithoutProducts#7 wRunOutBcd');
    AssertEquals_INT(Expected := 0, Actual := fbJamWithoutProducts.iCount, Message := 'JamWithoutProducts#7 iCount');
    AssertEquals_WORD(Expected := 16#0000,
                      Actual := fbJamWithoutProducts.wCountBcd,
                      Message := 'JamWithoutProducts#7 wCountBcd');

    // #8, t = 10500 мс — квитирование: затор снят
    GVL_S7Clock.tSimNow := T#10500MS;
    fbJamWithoutProducts.xAck := TRUE;
    fbJamWithoutProducts();
    AssertEquals_BOOL(Expected := FALSE, Actual := fbJamWithoutProducts.xHorn, Message := 'JamWithoutProducts#8 xHorn');
    AssertEquals_BOOL(Expected := FALSE,
                      Actual := fbJamWithoutProducts.xMotor,
                      Message := 'JamWithoutProducts#8 xMotor');
    AssertEquals_BOOL(Expected := FALSE,
                      Actual := fbJamWithoutProducts.xFlowOk,
                      Message := 'JamWithoutProducts#8 xFlowOk');
    AssertEquals_BOOL(Expected := FALSE, Actual := fbJamWithoutProducts.xJam, Message := 'JamWithoutProducts#8 xJam');
    AssertEquals_INT(Expected := 0,
                     Actual := fbJamWithoutProducts.iDelayLeft,
                     Message := 'JamWithoutProducts#8 iDelayLeft');
    AssertEquals_WORD(Expected := 16#0000,
                      Actual := fbJamWithoutProducts.wRunOutBcd,
                      Message := 'JamWithoutProducts#8 wRunOutBcd');
    AssertEquals_INT(Expected := 0, Actual := fbJamWithoutProducts.iCount, Message := 'JamWithoutProducts#8 iCount');
    AssertEquals_WORD(Expected := 16#0000,
                      Actual := fbJamWithoutProducts.wCountBcd,
                      Message := 'JamWithoutProducts#8 wCountBcd');

    // #9, t = 10600 мс — покой
    GVL_S7Clock.tSimNow := T#10600MS;
    fbJamWithoutProducts.xAck := FALSE;
    fbJamWithoutProducts();
    AssertEquals_BOOL(Expected := FALSE, Actual := fbJamWithoutProducts.xHorn, Message := 'JamWithoutProducts#9 xHorn');
    AssertEquals_BOOL(Expected := FALSE,
                      Actual := fbJamWithoutProducts.xMotor,
                      Message := 'JamWithoutProducts#9 xMotor');
    AssertEquals_BOOL(Expected := FALSE,
                      Actual := fbJamWithoutProducts.xFlowOk,
                      Message := 'JamWithoutProducts#9 xFlowOk');
    AssertEquals_BOOL(Expected := FALSE, Actual := fbJamWithoutProducts.xJam, Message := 'JamWithoutProducts#9 xJam');
    AssertEquals_INT(Expected := 0,
                     Actual := fbJamWithoutProducts.iDelayLeft,
                     Message := 'JamWithoutProducts#9 iDelayLeft');
    AssertEquals_WORD(Expected := 16#0000,
                      Actual := fbJamWithoutProducts.wRunOutBcd,
                      Message := 'JamWithoutProducts#9 wRunOutBcd');
    AssertEquals_INT(Expected := 0, Actual := fbJamWithoutProducts.iCount, Message := 'JamWithoutProducts#9 iCount');
    AssertEquals_WORD(Expected := 16#0000,
                      Actual := fbJamWithoutProducts.wCountBcd,
                      Message := 'JamWithoutProducts#9 wCountBcd');

    GVL_S7Clock.xSimulation := FALSE;
END_IF
coUnit.TEST_FINISHED();

(* ---- ProductsKeepFlow.method.decl.st ---- *)
// AUTO-GENERATED — не редактировать: scenarios/lang/FB_ConveyorStl.csv, сценарий ProductsKeepFlow (строк: 14)
METHOD PRIVATE ProductsKeepFlow
VAR
    stTimerZero : ST_S5Timer;  // пустое слово S5 для сброса
    stCounterZero : ST_S5Counter;  // пустое слово S5 для сброса
    iS5 : INT;  // номер таймера/счётчика S5
END_VAR

(* ---- ProductsKeepFlow.method.impl.st ---- *)
// AUTO-GENERATED — не редактировать: scenarios/lang/FB_ConveyorStl.csv, сценарий ProductsKeepFlow
coUnit.TEST('ProductsKeepFlow');
IF NOT xProductsKeepFlowDone THEN
    xProductsKeepFlowDone := TRUE;
    GVL_S7Clock.xSimulation := TRUE;
    // слова S5 — глобальные (GVL_S5Timers_Lang): сценарий начинается с чистых таймеров и счётчиков
    FOR iS5 := 0 TO 5 DO
        GVL_S5Timers_Lang.aTimer[iS5] := stTimerZero;
    END_FOR
    // слова S5 — глобальные (GVL_S5Counters_Lang): сценарий начинается с чистых таймеров и счётчиков
    FOR iS5 := 0 TO 1 DO
        GVL_S5Counters_Lang.aCounter[iS5] := stCounterZero;
    END_FOR

    // #1, t = 0 мс — пуск: запрос, сирена T1 и задержка T2 пошли
    GVL_S7Clock.tSimNow := T#0MS;
    fbProductsKeepFlow.xStart := TRUE;
    fbProductsKeepFlow.xStop := FALSE;
    fbProductsKeepFlow.xSensor := FALSE;
    fbProductsKeepFlow.xAck := FALSE;
    fbProductsKeepFlow.xCountReset := FALSE;
    fbProductsKeepFlow();
    AssertEquals_BOOL(Expected := TRUE, Actual := fbProductsKeepFlow.xHorn, Message := 'ProductsKeepFlow#1 xHorn');
    AssertEquals_BOOL(Expected := FALSE, Actual := fbProductsKeepFlow.xMotor, Message := 'ProductsKeepFlow#1 xMotor');
    AssertEquals_BOOL(Expected := FALSE, Actual := fbProductsKeepFlow.xFlowOk, Message := 'ProductsKeepFlow#1 xFlowOk');
    AssertEquals_BOOL(Expected := FALSE, Actual := fbProductsKeepFlow.xJam, Message := 'ProductsKeepFlow#1 xJam');
    AssertEquals_INT(Expected := 200,
                     Actual := fbProductsKeepFlow.iDelayLeft,
                     Message := 'ProductsKeepFlow#1 iDelayLeft');
    AssertEquals_WORD(Expected := 16#0000,
                      Actual := fbProductsKeepFlow.wRunOutBcd,
                      Message := 'ProductsKeepFlow#1 wRunOutBcd');
    AssertEquals_INT(Expected := 0, Actual := fbProductsKeepFlow.iCount, Message := 'ProductsKeepFlow#1 iCount');
    AssertEquals_WORD(Expected := 16#0000,
                      Actual := fbProductsKeepFlow.wCountBcd,
                      Message := 'ProductsKeepFlow#1 wCountBcd');

    // #2, t = 100 мс — кнопка отпущена
    GVL_S7Clock.tSimNow := T#100MS;
    fbProductsKeepFlow.xStart := FALSE;
    fbProductsKeepFlow();
    AssertEquals_BOOL(Expected := TRUE, Actual := fbProductsKeepFlow.xHorn, Message := 'ProductsKeepFlow#2 xHorn');
    AssertEquals_BOOL(Expected := FALSE, Actual := fbProductsKeepFlow.xMotor, Message := 'ProductsKeepFlow#2 xMotor');
    AssertEquals_BOOL(Expected := FALSE, Actual := fbProductsKeepFlow.xFlowOk, Message := 'ProductsKeepFlow#2 xFlowOk');
    AssertEquals_BOOL(Expected := FALSE, Actual := fbProductsKeepFlow.xJam, Message := 'ProductsKeepFlow#2 xJam');
    AssertEquals_INT(Expected := 190,
                     Actual := fbProductsKeepFlow.iDelayLeft,
                     Message := 'ProductsKeepFlow#2 iDelayLeft');
    AssertEquals_WORD(Expected := 16#0000,
                      Actual := fbProductsKeepFlow.wRunOutBcd,
                      Message := 'ProductsKeepFlow#2 wRunOutBcd');
    AssertEquals_INT(Expected := 0, Actual := fbProductsKeepFlow.iCount, Message := 'ProductsKeepFlow#2 iCount');
    AssertEquals_WORD(Expected := 16#0000,
                      Actual := fbProductsKeepFlow.wCountBcd,
                      Message := 'ProductsKeepFlow#2 wCountBcd');

    // #3, t = 2000 мс, на пороге таймера — 2 с: задержка T2 истекла — двигатель (T3 = 1)
    GVL_S7Clock.tSimNow := T#2000MS;
    fbProductsKeepFlow();
    AssertEquals_BOOL(Expected := FALSE, Actual := fbProductsKeepFlow.xHorn, Message := 'ProductsKeepFlow#3 xHorn');
    AssertEquals_BOOL(Expected := TRUE, Actual := fbProductsKeepFlow.xMotor, Message := 'ProductsKeepFlow#3 xMotor');
    AssertEquals_BOOL(Expected := FALSE, Actual := fbProductsKeepFlow.xFlowOk, Message := 'ProductsKeepFlow#3 xFlowOk');
    AssertEquals_BOOL(Expected := FALSE, Actual := fbProductsKeepFlow.xJam, Message := 'ProductsKeepFlow#3 xJam');
    AssertEquals_INT(Expected := 0,
                     Actual := fbProductsKeepFlow.iDelayLeft,
                     Message := 'ProductsKeepFlow#3 iDelayLeft');
    AssertEquals_WORD(Expected := 16#0000,
                      Actual := fbProductsKeepFlow.wRunOutBcd,
                      Message := 'ProductsKeepFlow#3 wRunOutBcd');
    AssertEquals_INT(Expected := 0, Actual := fbProductsKeepFlow.iCount, Message := 'ProductsKeepFlow#3 iCount');
    AssertEquals_WORD(Expected := 16#0000,
                      Actual := fbProductsKeepFlow.wCountBcd,
                      Message := 'ProductsKeepFlow#3 wCountBcd');

    // #4, t = 2500 мс — изделие №1: T4 пошёл
    GVL_S7Clock.tSimNow := T#2500MS;
    fbProductsKeepFlow.xSensor := TRUE;
    fbProductsKeepFlow();
    AssertEquals_BOOL(Expected := FALSE, Actual := fbProductsKeepFlow.xHorn, Message := 'ProductsKeepFlow#4 xHorn');
    AssertEquals_BOOL(Expected := TRUE, Actual := fbProductsKeepFlow.xMotor, Message := 'ProductsKeepFlow#4 xMotor');
    AssertEquals_BOOL(Expected := TRUE, Actual := fbProductsKeepFlow.xFlowOk, Message := 'ProductsKeepFlow#4 xFlowOk');
    AssertEquals_BOOL(Expected := FALSE, Actual := fbProductsKeepFlow.xJam, Message := 'ProductsKeepFlow#4 xJam');
    AssertEquals_INT(Expected := 0,
                     Actual := fbProductsKeepFlow.iDelayLeft,
                     Message := 'ProductsKeepFlow#4 iDelayLeft');
    AssertEquals_WORD(Expected := 16#0000,
                      Actual := fbProductsKeepFlow.wRunOutBcd,
                      Message := 'ProductsKeepFlow#4 wRunOutBcd');
    AssertEquals_INT(Expected := 1, Actual := fbProductsKeepFlow.iCount, Message := 'ProductsKeepFlow#4 iCount');
    AssertEquals_WORD(Expected := 16#0001,
                      Actual := fbProductsKeepFlow.wCountBcd,
                      Message := 'ProductsKeepFlow#4 wCountBcd');

    // #5, t = 2600 мс — датчик свободен
    GVL_S7Clock.tSimNow := T#2600MS;
    fbProductsKeepFlow.xSensor := FALSE;
    fbProductsKeepFlow();
    AssertEquals_BOOL(Expected := FALSE, Actual := fbProductsKeepFlow.xHorn, Message := 'ProductsKeepFlow#5 xHorn');
    AssertEquals_BOOL(Expected := TRUE, Actual := fbProductsKeepFlow.xMotor, Message := 'ProductsKeepFlow#5 xMotor');
    AssertEquals_BOOL(Expected := TRUE, Actual := fbProductsKeepFlow.xFlowOk, Message := 'ProductsKeepFlow#5 xFlowOk');
    AssertEquals_BOOL(Expected := FALSE, Actual := fbProductsKeepFlow.xJam, Message := 'ProductsKeepFlow#5 xJam');
    AssertEquals_INT(Expected := 0,
                     Actual := fbProductsKeepFlow.iDelayLeft,
                     Message := 'ProductsKeepFlow#5 iDelayLeft');
    AssertEquals_WORD(Expected := 16#0000,
                      Actual := fbProductsKeepFlow.wRunOutBcd,
                      Message := 'ProductsKeepFlow#5 wRunOutBcd');
    AssertEquals_INT(Expected := 1, Actual := fbProductsKeepFlow.iCount, Message := 'ProductsKeepFlow#5 iCount');
    AssertEquals_WORD(Expected := 16#0001,
                      Actual := fbProductsKeepFlow.wCountBcd,
                      Message := 'ProductsKeepFlow#5 wCountBcd');

    // #6, t = 4500 мс — изделие №2: T4 перезапущен
    GVL_S7Clock.tSimNow := T#4500MS;
    fbProductsKeepFlow.xSensor := TRUE;
    fbProductsKeepFlow();
    AssertEquals_BOOL(Expected := FALSE, Actual := fbProductsKeepFlow.xHorn, Message := 'ProductsKeepFlow#6 xHorn');
    AssertEquals_BOOL(Expected := TRUE, Actual := fbProductsKeepFlow.xMotor, Message := 'ProductsKeepFlow#6 xMotor');
    AssertEquals_BOOL(Expected := TRUE, Actual := fbProductsKeepFlow.xFlowOk, Message := 'ProductsKeepFlow#6 xFlowOk');
    AssertEquals_BOOL(Expected := FALSE, Actual := fbProductsKeepFlow.xJam, Message := 'ProductsKeepFlow#6 xJam');
    AssertEquals_INT(Expected := 0,
                     Actual := fbProductsKeepFlow.iDelayLeft,
                     Message := 'ProductsKeepFlow#6 iDelayLeft');
    AssertEquals_WORD(Expected := 16#0000,
                      Actual := fbProductsKeepFlow.wRunOutBcd,
                      Message := 'ProductsKeepFlow#6 wRunOutBcd');
    AssertEquals_INT(Expected := 2, Actual := fbProductsKeepFlow.iCount, Message := 'ProductsKeepFlow#6 iCount');
    AssertEquals_WORD(Expected := 16#0002,
                      Actual := fbProductsKeepFlow.wCountBcd,
                      Message := 'ProductsKeepFlow#6 wCountBcd');

    // #7, t = 4600 мс — датчик свободен
    GVL_S7Clock.tSimNow := T#4600MS;
    fbProductsKeepFlow.xSensor := FALSE;
    fbProductsKeepFlow();
    AssertEquals_BOOL(Expected := FALSE, Actual := fbProductsKeepFlow.xHorn, Message := 'ProductsKeepFlow#7 xHorn');
    AssertEquals_BOOL(Expected := TRUE, Actual := fbProductsKeepFlow.xMotor, Message := 'ProductsKeepFlow#7 xMotor');
    AssertEquals_BOOL(Expected := TRUE, Actual := fbProductsKeepFlow.xFlowOk, Message := 'ProductsKeepFlow#7 xFlowOk');
    AssertEquals_BOOL(Expected := FALSE, Actual := fbProductsKeepFlow.xJam, Message := 'ProductsKeepFlow#7 xJam');
    AssertEquals_INT(Expected := 0,
                     Actual := fbProductsKeepFlow.iDelayLeft,
                     Message := 'ProductsKeepFlow#7 iDelayLeft');
    AssertEquals_WORD(Expected := 16#0000,
                      Actual := fbProductsKeepFlow.wRunOutBcd,
                      Message := 'ProductsKeepFlow#7 wRunOutBcd');
    AssertEquals_INT(Expected := 2, Actual := fbProductsKeepFlow.iCount, Message := 'ProductsKeepFlow#7 iCount');
    AssertEquals_WORD(Expected := 16#0002,
                      Actual := fbProductsKeepFlow.wCountBcd,
                      Message := 'ProductsKeepFlow#7 wCountBcd');

    // #8, t = 6500 мс — изделие №3
    GVL_S7Clock.tSimNow := T#6500MS;
    fbProductsKeepFlow.xSensor := TRUE;
    fbProductsKeepFlow();
    AssertEquals_BOOL(Expected := FALSE, Actual := fbProductsKeepFlow.xHorn, Message := 'ProductsKeepFlow#8 xHorn');
    AssertEquals_BOOL(Expected := TRUE, Actual := fbProductsKeepFlow.xMotor, Message := 'ProductsKeepFlow#8 xMotor');
    AssertEquals_BOOL(Expected := TRUE, Actual := fbProductsKeepFlow.xFlowOk, Message := 'ProductsKeepFlow#8 xFlowOk');
    AssertEquals_BOOL(Expected := FALSE, Actual := fbProductsKeepFlow.xJam, Message := 'ProductsKeepFlow#8 xJam');
    AssertEquals_INT(Expected := 0,
                     Actual := fbProductsKeepFlow.iDelayLeft,
                     Message := 'ProductsKeepFlow#8 iDelayLeft');
    AssertEquals_WORD(Expected := 16#0000,
                      Actual := fbProductsKeepFlow.wRunOutBcd,
                      Message := 'ProductsKeepFlow#8 wRunOutBcd');
    AssertEquals_INT(Expected := 3, Actual := fbProductsKeepFlow.iCount, Message := 'ProductsKeepFlow#8 iCount');
    AssertEquals_WORD(Expected := 16#0003,
                      Actual := fbProductsKeepFlow.wCountBcd,
                      Message := 'ProductsKeepFlow#8 wCountBcd');

    // #9, t = 6600 мс — датчик свободен
    GVL_S7Clock.tSimNow := T#6600MS;
    fbProductsKeepFlow.xSensor := FALSE;
    fbProductsKeepFlow();
    AssertEquals_BOOL(Expected := FALSE, Actual := fbProductsKeepFlow.xHorn, Message := 'ProductsKeepFlow#9 xHorn');
    AssertEquals_BOOL(Expected := TRUE, Actual := fbProductsKeepFlow.xMotor, Message := 'ProductsKeepFlow#9 xMotor');
    AssertEquals_BOOL(Expected := TRUE, Actual := fbProductsKeepFlow.xFlowOk, Message := 'ProductsKeepFlow#9 xFlowOk');
    AssertEquals_BOOL(Expected := FALSE, Actual := fbProductsKeepFlow.xJam, Message := 'ProductsKeepFlow#9 xJam');
    AssertEquals_INT(Expected := 0,
                     Actual := fbProductsKeepFlow.iDelayLeft,
                     Message := 'ProductsKeepFlow#9 iDelayLeft');
    AssertEquals_WORD(Expected := 16#0000,
                      Actual := fbProductsKeepFlow.wRunOutBcd,
                      Message := 'ProductsKeepFlow#9 wRunOutBcd');
    AssertEquals_INT(Expected := 3, Actual := fbProductsKeepFlow.iCount, Message := 'ProductsKeepFlow#9 iCount');
    AssertEquals_WORD(Expected := 16#0003,
                      Actual := fbProductsKeepFlow.wCountBcd,
                      Message := 'ProductsKeepFlow#9 wCountBcd');

    // #10, t = 7000 мс, на пороге таймера — 5 с работы: контроль взведён, T4 идёт — затора нет
    GVL_S7Clock.tSimNow := T#7000MS;
    fbProductsKeepFlow();
    AssertEquals_BOOL(Expected := FALSE, Actual := fbProductsKeepFlow.xHorn, Message := 'ProductsKeepFlow#10 xHorn');
    AssertEquals_BOOL(Expected := TRUE, Actual := fbProductsKeepFlow.xMotor, Message := 'ProductsKeepFlow#10 xMotor');
    AssertEquals_BOOL(Expected := TRUE, Actual := fbProductsKeepFlow.xFlowOk, Message := 'ProductsKeepFlow#10 xFlowOk');
    AssertEquals_BOOL(Expected := FALSE, Actual := fbProductsKeepFlow.xJam, Message := 'ProductsKeepFlow#10 xJam');
    AssertEquals_INT(Expected := 0,
                     Actual := fbProductsKeepFlow.iDelayLeft,
                     Message := 'ProductsKeepFlow#10 iDelayLeft');
    AssertEquals_WORD(Expected := 16#0000,
                      Actual := fbProductsKeepFlow.wRunOutBcd,
                      Message := 'ProductsKeepFlow#10 wRunOutBcd');
    AssertEquals_INT(Expected := 3, Actual := fbProductsKeepFlow.iCount, Message := 'ProductsKeepFlow#10 iCount');
    AssertEquals_WORD(Expected := 16#0003,
                      Actual := fbProductsKeepFlow.wCountBcd,
                      Message := 'ProductsKeepFlow#10 wCountBcd');

    // #11, t = 8500 мс — изделие №4
    GVL_S7Clock.tSimNow := T#8500MS;
    fbProductsKeepFlow.xSensor := TRUE;
    fbProductsKeepFlow();
    AssertEquals_BOOL(Expected := FALSE, Actual := fbProductsKeepFlow.xHorn, Message := 'ProductsKeepFlow#11 xHorn');
    AssertEquals_BOOL(Expected := TRUE, Actual := fbProductsKeepFlow.xMotor, Message := 'ProductsKeepFlow#11 xMotor');
    AssertEquals_BOOL(Expected := TRUE, Actual := fbProductsKeepFlow.xFlowOk, Message := 'ProductsKeepFlow#11 xFlowOk');
    AssertEquals_BOOL(Expected := FALSE, Actual := fbProductsKeepFlow.xJam, Message := 'ProductsKeepFlow#11 xJam');
    AssertEquals_INT(Expected := 0,
                     Actual := fbProductsKeepFlow.iDelayLeft,
                     Message := 'ProductsKeepFlow#11 iDelayLeft');
    AssertEquals_WORD(Expected := 16#0000,
                      Actual := fbProductsKeepFlow.wRunOutBcd,
                      Message := 'ProductsKeepFlow#11 wRunOutBcd');
    AssertEquals_INT(Expected := 4, Actual := fbProductsKeepFlow.iCount, Message := 'ProductsKeepFlow#11 iCount');
    AssertEquals_WORD(Expected := 16#0004,
                      Actual := fbProductsKeepFlow.wCountBcd,
                      Message := 'ProductsKeepFlow#11 wCountBcd');

    // #12, t = 8600 мс — датчик свободен
    GVL_S7Clock.tSimNow := T#8600MS;
    fbProductsKeepFlow.xSensor := FALSE;
    fbProductsKeepFlow();
    AssertEquals_BOOL(Expected := FALSE, Actual := fbProductsKeepFlow.xHorn, Message := 'ProductsKeepFlow#12 xHorn');
    AssertEquals_BOOL(Expected := TRUE, Actual := fbProductsKeepFlow.xMotor, Message := 'ProductsKeepFlow#12 xMotor');
    AssertEquals_BOOL(Expected := TRUE, Actual := fbProductsKeepFlow.xFlowOk, Message := 'ProductsKeepFlow#12 xFlowOk');
    AssertEquals_BOOL(Expected := FALSE, Actual := fbProductsKeepFlow.xJam, Message := 'ProductsKeepFlow#12 xJam');
    AssertEquals_INT(Expected := 0,
                     Actual := fbProductsKeepFlow.iDelayLeft,
                     Message := 'ProductsKeepFlow#12 iDelayLeft');
    AssertEquals_WORD(Expected := 16#0000,
                      Actual := fbProductsKeepFlow.wRunOutBcd,
                      Message := 'ProductsKeepFlow#12 wRunOutBcd');
    AssertEquals_INT(Expected := 4, Actual := fbProductsKeepFlow.iCount, Message := 'ProductsKeepFlow#12 iCount');
    AssertEquals_WORD(Expected := 16#0004,
                      Actual := fbProductsKeepFlow.wCountBcd,
                      Message := 'ProductsKeepFlow#12 wCountBcd');

    // #13, t = 10600 мс — 2,1 с без изделий
    GVL_S7Clock.tSimNow := T#10600MS;
    fbProductsKeepFlow();
    AssertEquals_BOOL(Expected := FALSE, Actual := fbProductsKeepFlow.xHorn, Message := 'ProductsKeepFlow#13 xHorn');
    AssertEquals_BOOL(Expected := TRUE, Actual := fbProductsKeepFlow.xMotor, Message := 'ProductsKeepFlow#13 xMotor');
    AssertEquals_BOOL(Expected := TRUE, Actual := fbProductsKeepFlow.xFlowOk, Message := 'ProductsKeepFlow#13 xFlowOk');
    AssertEquals_BOOL(Expected := FALSE, Actual := fbProductsKeepFlow.xJam, Message := 'ProductsKeepFlow#13 xJam');
    AssertEquals_INT(Expected := 0,
                     Actual := fbProductsKeepFlow.iDelayLeft,
                     Message := 'ProductsKeepFlow#13 iDelayLeft');
    AssertEquals_WORD(Expected := 16#0000,
                      Actual := fbProductsKeepFlow.wRunOutBcd,
                      Message := 'ProductsKeepFlow#13 wRunOutBcd');
    AssertEquals_INT(Expected := 4, Actual := fbProductsKeepFlow.iCount, Message := 'ProductsKeepFlow#13 iCount');
    AssertEquals_WORD(Expected := 16#0004,
                      Actual := fbProductsKeepFlow.wCountBcd,
                      Message := 'ProductsKeepFlow#13 wCountBcd');

    // #14, t = 12500 мс, на пороге таймера — 4 с без изделий: T4 истёк — затор
    GVL_S7Clock.tSimNow := T#12500MS;
    fbProductsKeepFlow();
    AssertEquals_BOOL(Expected := FALSE, Actual := fbProductsKeepFlow.xHorn, Message := 'ProductsKeepFlow#14 xHorn');
    AssertEquals_BOOL(Expected := TRUE, Actual := fbProductsKeepFlow.xMotor, Message := 'ProductsKeepFlow#14 xMotor');
    AssertEquals_BOOL(Expected := FALSE,
                      Actual := fbProductsKeepFlow.xFlowOk,
                      Message := 'ProductsKeepFlow#14 xFlowOk');
    AssertEquals_BOOL(Expected := TRUE, Actual := fbProductsKeepFlow.xJam, Message := 'ProductsKeepFlow#14 xJam');
    AssertEquals_INT(Expected := 0,
                     Actual := fbProductsKeepFlow.iDelayLeft,
                     Message := 'ProductsKeepFlow#14 iDelayLeft');
    AssertEquals_WORD(Expected := 16#0000,
                      Actual := fbProductsKeepFlow.wRunOutBcd,
                      Message := 'ProductsKeepFlow#14 wRunOutBcd');
    AssertEquals_INT(Expected := 4, Actual := fbProductsKeepFlow.iCount, Message := 'ProductsKeepFlow#14 iCount');
    AssertEquals_WORD(Expected := 16#0004,
                      Actual := fbProductsKeepFlow.wCountBcd,
                      Message := 'ProductsKeepFlow#14 wCountBcd');

    GVL_S7Clock.xSimulation := FALSE;
END_IF
coUnit.TEST_FINISHED();

(* ---- StartSequence.method.decl.st ---- *)
// AUTO-GENERATED — не редактировать: scenarios/lang/FB_ConveyorStl.csv, сценарий StartSequence (строк: 6)
METHOD PRIVATE StartSequence
VAR
    stTimerZero : ST_S5Timer;  // пустое слово S5 для сброса
    stCounterZero : ST_S5Counter;  // пустое слово S5 для сброса
    iS5 : INT;  // номер таймера/счётчика S5
END_VAR

(* ---- StartSequence.method.impl.st ---- *)
// AUTO-GENERATED — не редактировать: scenarios/lang/FB_ConveyorStl.csv, сценарий StartSequence
coUnit.TEST('StartSequence');
IF NOT xStartSequenceDone THEN
    xStartSequenceDone := TRUE;
    GVL_S7Clock.xSimulation := TRUE;
    // слова S5 — глобальные (GVL_S5Timers_Lang): сценарий начинается с чистых таймеров и счётчиков
    FOR iS5 := 0 TO 5 DO
        GVL_S5Timers_Lang.aTimer[iS5] := stTimerZero;
    END_FOR
    // слова S5 — глобальные (GVL_S5Counters_Lang): сценарий начинается с чистых таймеров и счётчиков
    FOR iS5 := 0 TO 1 DO
        GVL_S5Counters_Lang.aCounter[iS5] := stCounterZero;
    END_FOR

    // #1, t = 0 мс — пуск: сирена и задержка, остаток 200 единиц
    GVL_S7Clock.tSimNow := T#0MS;
    fbStartSequence.xStart := TRUE;
    fbStartSequence.xStop := FALSE;
    fbStartSequence.xSensor := FALSE;
    fbStartSequence.xAck := FALSE;
    fbStartSequence.xCountReset := FALSE;
    fbStartSequence();
    AssertEquals_BOOL(Expected := TRUE, Actual := fbStartSequence.xHorn, Message := 'StartSequence#1 xHorn');
    AssertEquals_BOOL(Expected := FALSE, Actual := fbStartSequence.xMotor, Message := 'StartSequence#1 xMotor');
    AssertEquals_BOOL(Expected := FALSE, Actual := fbStartSequence.xFlowOk, Message := 'StartSequence#1 xFlowOk');
    AssertEquals_BOOL(Expected := FALSE, Actual := fbStartSequence.xJam, Message := 'StartSequence#1 xJam');
    AssertEquals_INT(Expected := 200, Actual := fbStartSequence.iDelayLeft, Message := 'StartSequence#1 iDelayLeft');
    AssertEquals_WORD(Expected := 16#0000,
                      Actual := fbStartSequence.wRunOutBcd,
                      Message := 'StartSequence#1 wRunOutBcd');
    AssertEquals_INT(Expected := 0, Actual := fbStartSequence.iCount, Message := 'StartSequence#1 iCount');
    AssertEquals_WORD(Expected := 16#0000, Actual := fbStartSequence.wCountBcd, Message := 'StartSequence#1 wCountBcd');

    // #2, t = 300 мс — кнопка отпущена: сирена звучит, остаток 170
    GVL_S7Clock.tSimNow := T#300MS;
    fbStartSequence.xStart := FALSE;
    fbStartSequence();
    AssertEquals_BOOL(Expected := TRUE, Actual := fbStartSequence.xHorn, Message := 'StartSequence#2 xHorn');
    AssertEquals_BOOL(Expected := FALSE, Actual := fbStartSequence.xMotor, Message := 'StartSequence#2 xMotor');
    AssertEquals_BOOL(Expected := FALSE, Actual := fbStartSequence.xFlowOk, Message := 'StartSequence#2 xFlowOk');
    AssertEquals_BOOL(Expected := FALSE, Actual := fbStartSequence.xJam, Message := 'StartSequence#2 xJam');
    AssertEquals_INT(Expected := 170, Actual := fbStartSequence.iDelayLeft, Message := 'StartSequence#2 iDelayLeft');
    AssertEquals_WORD(Expected := 16#0000,
                      Actual := fbStartSequence.wRunOutBcd,
                      Message := 'StartSequence#2 wRunOutBcd');
    AssertEquals_INT(Expected := 0, Actual := fbStartSequence.iCount, Message := 'StartSequence#2 iCount');
    AssertEquals_WORD(Expected := 16#0000, Actual := fbStartSequence.wCountBcd, Message := 'StartSequence#2 wCountBcd');

    // #3, t = 1000 мс, на пороге таймера — 1 с: сирена выключилась (T1 истёк), остаток 100
    GVL_S7Clock.tSimNow := T#1000MS;
    fbStartSequence();
    AssertEquals_BOOL(Expected := FALSE, Actual := fbStartSequence.xHorn, Message := 'StartSequence#3 xHorn');
    AssertEquals_BOOL(Expected := FALSE, Actual := fbStartSequence.xMotor, Message := 'StartSequence#3 xMotor');
    AssertEquals_BOOL(Expected := FALSE, Actual := fbStartSequence.xFlowOk, Message := 'StartSequence#3 xFlowOk');
    AssertEquals_BOOL(Expected := FALSE, Actual := fbStartSequence.xJam, Message := 'StartSequence#3 xJam');
    AssertEquals_INT(Expected := 100, Actual := fbStartSequence.iDelayLeft, Message := 'StartSequence#3 iDelayLeft');
    AssertEquals_WORD(Expected := 16#0000,
                      Actual := fbStartSequence.wRunOutBcd,
                      Message := 'StartSequence#3 wRunOutBcd');
    AssertEquals_INT(Expected := 0, Actual := fbStartSequence.iCount, Message := 'StartSequence#3 iCount');
    AssertEquals_WORD(Expected := 16#0000, Actual := fbStartSequence.wCountBcd, Message := 'StartSequence#3 wCountBcd');

    // #4, t = 1500 мс — остаток 50
    GVL_S7Clock.tSimNow := T#1500MS;
    fbStartSequence();
    AssertEquals_BOOL(Expected := FALSE, Actual := fbStartSequence.xHorn, Message := 'StartSequence#4 xHorn');
    AssertEquals_BOOL(Expected := FALSE, Actual := fbStartSequence.xMotor, Message := 'StartSequence#4 xMotor');
    AssertEquals_BOOL(Expected := FALSE, Actual := fbStartSequence.xFlowOk, Message := 'StartSequence#4 xFlowOk');
    AssertEquals_BOOL(Expected := FALSE, Actual := fbStartSequence.xJam, Message := 'StartSequence#4 xJam');
    AssertEquals_INT(Expected := 50, Actual := fbStartSequence.iDelayLeft, Message := 'StartSequence#4 iDelayLeft');
    AssertEquals_WORD(Expected := 16#0000,
                      Actual := fbStartSequence.wRunOutBcd,
                      Message := 'StartSequence#4 wRunOutBcd');
    AssertEquals_INT(Expected := 0, Actual := fbStartSequence.iCount, Message := 'StartSequence#4 iCount');
    AssertEquals_WORD(Expected := 16#0000, Actual := fbStartSequence.wCountBcd, Message := 'StartSequence#4 wCountBcd');

    // #5, t = 2000 мс, на пороге таймера — 2 с: задержка истекла — двигатель
    GVL_S7Clock.tSimNow := T#2000MS;
    fbStartSequence();
    AssertEquals_BOOL(Expected := FALSE, Actual := fbStartSequence.xHorn, Message := 'StartSequence#5 xHorn');
    AssertEquals_BOOL(Expected := TRUE, Actual := fbStartSequence.xMotor, Message := 'StartSequence#5 xMotor');
    AssertEquals_BOOL(Expected := FALSE, Actual := fbStartSequence.xFlowOk, Message := 'StartSequence#5 xFlowOk');
    AssertEquals_BOOL(Expected := FALSE, Actual := fbStartSequence.xJam, Message := 'StartSequence#5 xJam');
    AssertEquals_INT(Expected := 0, Actual := fbStartSequence.iDelayLeft, Message := 'StartSequence#5 iDelayLeft');
    AssertEquals_WORD(Expected := 16#0000,
                      Actual := fbStartSequence.wRunOutBcd,
                      Message := 'StartSequence#5 wRunOutBcd');
    AssertEquals_INT(Expected := 0, Actual := fbStartSequence.iCount, Message := 'StartSequence#5 iCount');
    AssertEquals_WORD(Expected := 16#0000, Actual := fbStartSequence.wCountBcd, Message := 'StartSequence#5 wCountBcd');

    // #6, t = 2500 мс — работает
    GVL_S7Clock.tSimNow := T#2500MS;
    fbStartSequence();
    AssertEquals_BOOL(Expected := FALSE, Actual := fbStartSequence.xHorn, Message := 'StartSequence#6 xHorn');
    AssertEquals_BOOL(Expected := TRUE, Actual := fbStartSequence.xMotor, Message := 'StartSequence#6 xMotor');
    AssertEquals_BOOL(Expected := FALSE, Actual := fbStartSequence.xFlowOk, Message := 'StartSequence#6 xFlowOk');
    AssertEquals_BOOL(Expected := FALSE, Actual := fbStartSequence.xJam, Message := 'StartSequence#6 xJam');
    AssertEquals_INT(Expected := 0, Actual := fbStartSequence.iDelayLeft, Message := 'StartSequence#6 iDelayLeft');
    AssertEquals_WORD(Expected := 16#0000,
                      Actual := fbStartSequence.wRunOutBcd,
                      Message := 'StartSequence#6 wRunOutBcd');
    AssertEquals_INT(Expected := 0, Actual := fbStartSequence.iCount, Message := 'StartSequence#6 iCount');
    AssertEquals_WORD(Expected := 16#0000, Actual := fbStartSequence.wCountBcd, Message := 'StartSequence#6 wCountBcd');

    GVL_S7Clock.xSimulation := FALSE;
END_IF
coUnit.TEST_FINISHED();

(* ---- StopRunOut.method.decl.st ---- *)
// AUTO-GENERATED — не редактировать: scenarios/lang/FB_ConveyorStl.csv, сценарий StopRunOut (строк: 7)
METHOD PRIVATE StopRunOut
VAR
    stTimerZero : ST_S5Timer;  // пустое слово S5 для сброса
    stCounterZero : ST_S5Counter;  // пустое слово S5 для сброса
    iS5 : INT;  // номер таймера/счётчика S5
END_VAR

(* ---- StopRunOut.method.impl.st ---- *)
// AUTO-GENERATED — не редактировать: scenarios/lang/FB_ConveyorStl.csv, сценарий StopRunOut
coUnit.TEST('StopRunOut');
IF NOT xStopRunOutDone THEN
    xStopRunOutDone := TRUE;
    GVL_S7Clock.xSimulation := TRUE;
    // слова S5 — глобальные (GVL_S5Timers_Lang): сценарий начинается с чистых таймеров и счётчиков
    FOR iS5 := 0 TO 5 DO
        GVL_S5Timers_Lang.aTimer[iS5] := stTimerZero;
    END_FOR
    // слова S5 — глобальные (GVL_S5Counters_Lang): сценарий начинается с чистых таймеров и счётчиков
    FOR iS5 := 0 TO 1 DO
        GVL_S5Counters_Lang.aCounter[iS5] := stCounterZero;
    END_FOR

    // #1, t = 0 мс — пуск: запрос, сирена T1 и задержка T2 пошли
    GVL_S7Clock.tSimNow := T#0MS;
    fbStopRunOut.xStart := TRUE;
    fbStopRunOut.xStop := FALSE;
    fbStopRunOut.xSensor := FALSE;
    fbStopRunOut.xAck := FALSE;
    fbStopRunOut.xCountReset := FALSE;
    fbStopRunOut();
    AssertEquals_BOOL(Expected := TRUE, Actual := fbStopRunOut.xHorn, Message := 'StopRunOut#1 xHorn');
    AssertEquals_BOOL(Expected := FALSE, Actual := fbStopRunOut.xMotor, Message := 'StopRunOut#1 xMotor');
    AssertEquals_BOOL(Expected := FALSE, Actual := fbStopRunOut.xFlowOk, Message := 'StopRunOut#1 xFlowOk');
    AssertEquals_BOOL(Expected := FALSE, Actual := fbStopRunOut.xJam, Message := 'StopRunOut#1 xJam');
    AssertEquals_INT(Expected := 200, Actual := fbStopRunOut.iDelayLeft, Message := 'StopRunOut#1 iDelayLeft');
    AssertEquals_WORD(Expected := 16#0000, Actual := fbStopRunOut.wRunOutBcd, Message := 'StopRunOut#1 wRunOutBcd');
    AssertEquals_INT(Expected := 0, Actual := fbStopRunOut.iCount, Message := 'StopRunOut#1 iCount');
    AssertEquals_WORD(Expected := 16#0000, Actual := fbStopRunOut.wCountBcd, Message := 'StopRunOut#1 wCountBcd');

    // #2, t = 100 мс — кнопка отпущена
    GVL_S7Clock.tSimNow := T#100MS;
    fbStopRunOut.xStart := FALSE;
    fbStopRunOut();
    AssertEquals_BOOL(Expected := TRUE, Actual := fbStopRunOut.xHorn, Message := 'StopRunOut#2 xHorn');
    AssertEquals_BOOL(Expected := FALSE, Actual := fbStopRunOut.xMotor, Message := 'StopRunOut#2 xMotor');
    AssertEquals_BOOL(Expected := FALSE, Actual := fbStopRunOut.xFlowOk, Message := 'StopRunOut#2 xFlowOk');
    AssertEquals_BOOL(Expected := FALSE, Actual := fbStopRunOut.xJam, Message := 'StopRunOut#2 xJam');
    AssertEquals_INT(Expected := 190, Actual := fbStopRunOut.iDelayLeft, Message := 'StopRunOut#2 iDelayLeft');
    AssertEquals_WORD(Expected := 16#0000, Actual := fbStopRunOut.wRunOutBcd, Message := 'StopRunOut#2 wRunOutBcd');
    AssertEquals_INT(Expected := 0, Actual := fbStopRunOut.iCount, Message := 'StopRunOut#2 iCount');
    AssertEquals_WORD(Expected := 16#0000, Actual := fbStopRunOut.wCountBcd, Message := 'StopRunOut#2 wCountBcd');

    // #3, t = 2000 мс, на пороге таймера — 2 с: задержка T2 истекла — двигатель (T3 = 1)
    GVL_S7Clock.tSimNow := T#2000MS;
    fbStopRunOut();
    AssertEquals_BOOL(Expected := FALSE, Actual := fbStopRunOut.xHorn, Message := 'StopRunOut#3 xHorn');
    AssertEquals_BOOL(Expected := TRUE, Actual := fbStopRunOut.xMotor, Message := 'StopRunOut#3 xMotor');
    AssertEquals_BOOL(Expected := FALSE, Actual := fbStopRunOut.xFlowOk, Message := 'StopRunOut#3 xFlowOk');
    AssertEquals_BOOL(Expected := FALSE, Actual := fbStopRunOut.xJam, Message := 'StopRunOut#3 xJam');
    AssertEquals_INT(Expected := 0, Actual := fbStopRunOut.iDelayLeft, Message := 'StopRunOut#3 iDelayLeft');
    AssertEquals_WORD(Expected := 16#0000, Actual := fbStopRunOut.wRunOutBcd, Message := 'StopRunOut#3 wRunOutBcd');
    AssertEquals_INT(Expected := 0, Actual := fbStopRunOut.iCount, Message := 'StopRunOut#3 iCount');
    AssertEquals_WORD(Expected := 16#0000, Actual := fbStopRunOut.wCountBcd, Message := 'StopRunOut#3 wCountBcd');

    // #4, t = 3000 мс — стоп: запрос снят, выбег T3 пошёл, 16#0300
    GVL_S7Clock.tSimNow := T#3000MS;
    fbStopRunOut.xStop := TRUE;
    fbStopRunOut();
    AssertEquals_BOOL(Expected := FALSE, Actual := fbStopRunOut.xHorn, Message := 'StopRunOut#4 xHorn');
    AssertEquals_BOOL(Expected := TRUE, Actual := fbStopRunOut.xMotor, Message := 'StopRunOut#4 xMotor');
    AssertEquals_BOOL(Expected := FALSE, Actual := fbStopRunOut.xFlowOk, Message := 'StopRunOut#4 xFlowOk');
    AssertEquals_BOOL(Expected := FALSE, Actual := fbStopRunOut.xJam, Message := 'StopRunOut#4 xJam');
    AssertEquals_INT(Expected := 0, Actual := fbStopRunOut.iDelayLeft, Message := 'StopRunOut#4 iDelayLeft');
    AssertEquals_WORD(Expected := 16#0300, Actual := fbStopRunOut.wRunOutBcd, Message := 'StopRunOut#4 wRunOutBcd');
    AssertEquals_INT(Expected := 0, Actual := fbStopRunOut.iCount, Message := 'StopRunOut#4 iCount');
    AssertEquals_WORD(Expected := 16#0000, Actual := fbStopRunOut.wCountBcd, Message := 'StopRunOut#4 wCountBcd');

    // #5, t = 3100 мс — выбег: остаток 290 единиц
    GVL_S7Clock.tSimNow := T#3100MS;
    fbStopRunOut.xStop := FALSE;
    fbStopRunOut();
    AssertEquals_BOOL(Expected := FALSE, Actual := fbStopRunOut.xHorn, Message := 'StopRunOut#5 xHorn');
    AssertEquals_BOOL(Expected := TRUE, Actual := fbStopRunOut.xMotor, Message := 'StopRunOut#5 xMotor');
    AssertEquals_BOOL(Expected := FALSE, Actual := fbStopRunOut.xFlowOk, Message := 'StopRunOut#5 xFlowOk');
    AssertEquals_BOOL(Expected := FALSE, Actual := fbStopRunOut.xJam, Message := 'StopRunOut#5 xJam');
    AssertEquals_INT(Expected := 0, Actual := fbStopRunOut.iDelayLeft, Message := 'StopRunOut#5 iDelayLeft');
    AssertEquals_WORD(Expected := 16#0290, Actual := fbStopRunOut.wRunOutBcd, Message := 'StopRunOut#5 wRunOutBcd');
    AssertEquals_INT(Expected := 0, Actual := fbStopRunOut.iCount, Message := 'StopRunOut#5 iCount');
    AssertEquals_WORD(Expected := 16#0000, Actual := fbStopRunOut.wCountBcd, Message := 'StopRunOut#5 wCountBcd');

    // #6, t = 4500 мс — выбег: остаток 150 единиц
    GVL_S7Clock.tSimNow := T#4500MS;
    fbStopRunOut();
    AssertEquals_BOOL(Expected := FALSE, Actual := fbStopRunOut.xHorn, Message := 'StopRunOut#6 xHorn');
    AssertEquals_BOOL(Expected := TRUE, Actual := fbStopRunOut.xMotor, Message := 'StopRunOut#6 xMotor');
    AssertEquals_BOOL(Expected := FALSE, Actual := fbStopRunOut.xFlowOk, Message := 'StopRunOut#6 xFlowOk');
    AssertEquals_BOOL(Expected := FALSE, Actual := fbStopRunOut.xJam, Message := 'StopRunOut#6 xJam');
    AssertEquals_INT(Expected := 0, Actual := fbStopRunOut.iDelayLeft, Message := 'StopRunOut#6 iDelayLeft');
    AssertEquals_WORD(Expected := 16#0150, Actual := fbStopRunOut.wRunOutBcd, Message := 'StopRunOut#6 wRunOutBcd');
    AssertEquals_INT(Expected := 0, Actual := fbStopRunOut.iCount, Message := 'StopRunOut#6 iCount');
    AssertEquals_WORD(Expected := 16#0000, Actual := fbStopRunOut.wCountBcd, Message := 'StopRunOut#6 wCountBcd');

    // #7, t = 6000 мс, на пороге таймера — 3 с выбега: двигатель остановлен
    GVL_S7Clock.tSimNow := T#6000MS;
    fbStopRunOut();
    AssertEquals_BOOL(Expected := FALSE, Actual := fbStopRunOut.xHorn, Message := 'StopRunOut#7 xHorn');
    AssertEquals_BOOL(Expected := FALSE, Actual := fbStopRunOut.xMotor, Message := 'StopRunOut#7 xMotor');
    AssertEquals_BOOL(Expected := FALSE, Actual := fbStopRunOut.xFlowOk, Message := 'StopRunOut#7 xFlowOk');
    AssertEquals_BOOL(Expected := FALSE, Actual := fbStopRunOut.xJam, Message := 'StopRunOut#7 xJam');
    AssertEquals_INT(Expected := 0, Actual := fbStopRunOut.iDelayLeft, Message := 'StopRunOut#7 iDelayLeft');
    AssertEquals_WORD(Expected := 16#0000, Actual := fbStopRunOut.wRunOutBcd, Message := 'StopRunOut#7 wRunOutBcd');
    AssertEquals_INT(Expected := 0, Actual := fbStopRunOut.iCount, Message := 'StopRunOut#7 iCount');
    AssertEquals_WORD(Expected := 16#0000, Actual := fbStopRunOut.wCountBcd, Message := 'StopRunOut#7 wCountBcd');

    GVL_S7Clock.xSimulation := FALSE;
END_IF
coUnit.TEST_FINISHED();
